(* IEC 61131-3 sources: plc-st-coding-agent/progress/evidence/f14_v14_remaining_20261113/jobs/custom_minimax-m27 (part 6) *)

(* ---- public-medium-06.raw_candidate_02.st ---- *)
FUNCTION_BLOCK FB_SlabThicknessMonitor
(*
 * ENGINEERING_CONTRACT
 * =============================================================================
 * Output/State          | Activation          | Retention            | Reset/Deactivation            | Units
 * ----------------------+---------------------+----------------------+-------------------------------+-----------------
 * THICKNESS_ALARM       | Rising edge valid   | Min 500ms hold;      | Signal invalid clears all     | BOOL
 *                       | THICKNESS_FAULT     | continues if fault   | alarm and hold state (PUB001) |
 * Alarm hold timer      | TON(IN: valid &     | TON.ET saturates at  | Signal invalid resets TON     | LTIME (≥500ms)
 *                       |   (fault OR holding))| PT=500ms            |                               |
 * Holding flag          | Fault OR holding    | Self-holds while     | Signal invalid clears         | BOOL
 *                       |                     |   fault OR timer run |                               |
 * Slab_Fault_Counter    | FALSE→TRUE valid    | Accumulates monoton  | None by task spec             | UINT
 *                       | fault transition    | (never auto-reset)   |                               |
 * Slab_Fault_History[0] | New fault entry     | Shifts [n]→[n+1]     | Power-up init to 0            | ARRAY[0..4] DINT
 *                       | writes to index 0   | (0 newest)           |                               |
 * Slab_Runtime_Accumulator| While CUTTING_RUN  | Preserved when       | None by task spec             | LTIME (accumulates)
 *                       | + valid + no fault  | conditions not met   |                               |
 * =============================================================================
 * CONTRACT_RULES [{"kind": "hold_until_reset", "output": "THICKNESS_ALARM", "set_input": "THICKNESS_FAULT", "reset_input": null}]
 *)

VAR_INPUT
    THICKNESS_FAULT        : BOOL;
    THICKNESS_SIGNAL_VALID : BOOL;
    CUTTING_RUN            : BOOL;
    FaultTimestamp         : DINT;
    CycleTime              : TIME;
END_VAR

VAR_OUTPUT
    THICKNESS_ALARM           : BOOL;
    Slab_Fault_Counter        : UINT;
    Slab_Runtime_Accumulator  : LTIME;
    Slab_Fault_History        : ARRAY[0..4] OF DINT;
END_VAR

VAR
    faultRisingEdge    : R_TRIG;
    signalValidPrev    : BOOL;
    alarmHoldTimer     : TON;
    alarmHolding       : BOOL;
    faultActive        : BOOL;
END_VAR

// ---------------------------------------------------------------------------
// Power-up initialization (first scan after instantiation)
// ---------------------------------------------------------------------------
IF NOT alarmHoldTimer.Q AND NOT faultActive AND NOT alarmHolding THEN
    Slab_Fault_Counter       := 0;
    Slab_Runtime_Accumulator := LTIME#0;
    Slab_Fault_History[0]    := 0;
    Slab_Fault_History[1]    := 0;
    Slab_Fault_History[2]    := 0;
    Slab_Fault_History[3]    := 0;
    Slab_Fault_History[4]    := 0;
END_IF;

// ---------------------------------------------------------------------------
// Detect FALSE→TRUE transition on valid fault signal
// ---------------------------------------------------------------------------
faultRisingEdge(CLK := THICKNESS_FAULT AND THICKNESS_SIGNAL_VALID);

// ---------------------------------------------------------------------------
// Handle signal-valid transitions: clear alarm/hold when signal lost (PUB001)
// ---------------------------------------------------------------------------
IF THICKNESS_SIGNAL_VALID THEN
    IF NOT signalValidPrev THEN
        // Signal just restored after being invalid
        alarmHolding  := FALSE;
        alarmHoldTimer(IN := FALSE);
        faultActive   := FALSE;
    END_IF;

    // -------------------------------------------------------------------------
    // On rising edge of valid fault: record entry and start hold
    // -------------------------------------------------------------------------
    IF faultRisingEdge.Q THEN
        // Increment counter
        Slab_Fault_Counter := Slab_Fault_Counter + UINT#1;

        // Shift history: index 3→4, 2→3, 1→2, 0→1, then write new to 0
        Slab_Fault_History[4] := Slab_Fault_History[3];
        Slab_Fault_History[3] := Slab_Fault_History[2];
        Slab_Fault_History[2] := Slab_Fault_History[1];
        Slab_Fault_History[1] := Slab_Fault_History[0];
        Slab_Fault_History[0] := FaultTimestamp;

        // Activate alarm and start 500 ms hold timer
        faultActive        := TRUE;
        alarmHolding       := TRUE;
        alarmHoldTimer(IN  := TRUE, PT := T#500ms);
    END_IF;

    // -------------------------------------------------------------------------
    // Update alarm state: hold while fault persists or timer running
    // -------------------------------------------------------------------------
    IF faultActive THEN
        // Keep timer running while fault is present
        alarmHoldTimer(IN := TRUE, PT := T#500ms);

        // Alarm stays active while fault or hold timer active
        alarmHolding := THICKNESS_FAULT OR alarmHoldTimer.Q;

        // Release hold tracking once fault clears and timer completes
        IF NOT THICKNESS_FAULT AND alarmHolding AND NOT alarmHoldTimer.Q THEN
            alarmHolding := FALSE;
        END_IF;

        // Clear fault-active flag when fault goes away (hold may continue)
        IF NOT THICKNESS_FAULT THEN
            faultActive := FALSE;
        END_IF;
    END_IF;

    // Final alarm output
    THICKNESS_ALARM := alarmHolding OR faultActive;

    // -------------------------------------------------------------------------
    // Runtime accumulation: only while cutting, signal valid, no fault
    // -------------------------------------------------------------------------
    IF CUTTING_RUN AND NOT THICKNESS_FAULT THEN
        Slab_Runtime_Accumulator := Slab_Runtime_Accumulator + TO_LTIME(CycleTime);
    END_IF;

ELSE
    // Signal invalid: clear alarm and all hold state (PUB001)
    THICKNESS_ALARM  := FALSE;
    alarmHolding     := FALSE;
    faultActive      := FALSE;
    alarmHoldTimer(IN := FALSE);
END_IF;

// ---------------------------------------------------------------------------
// Latch previous scan signal-valid state for edge detection
// ---------------------------------------------------------------------------
signalValidPrev := THICKNESS_SIGNAL_VALID;

END_FUNCTION_BLOCK

(* ---- public-medium-06.raw_candidate_03.st ---- *)
FUNCTION_BLOCK FB_SlabThicknessMonitor
(*
 * ENGINEERING_CONTRACT
 * =============================================================================
 * Output/State          | Activation          | Retention            | Reset/Deactivation            | Units
 * ----------------------+---------------------+----------------------+-------------------------------+-----------------
 * THICKNESS_ALARM       | Rising edge valid   | Min 500ms hold;      | Signal invalid clears all     | BOOL
 *                       | THICKNESS_FAULT     | continues if fault   | alarm and hold state (PUB001) |
 * Alarm hold timer      | TON(IN: valid &     | TON.ET saturates at  | Signal invalid resets TON     | LTIME (≥500ms)
 *                       |   (fault OR holding))| PT=500ms            |                               |
 * Holding flag          | Fault OR holding    | Self-holds while     | Signal invalid clears         | BOOL
 *                       |                     |   fault OR timer run |                               |
 * Slab_Fault_Counter    | FALSE→TRUE valid    | Accumulates monoton  | None by task spec             | UINT
 *                       | fault transition    | (never auto-reset)   |                               |
 * Slab_Fault_History[0] | New fault entry     | Shifts [n]→[n+1]     | Power-up init to 0            | ARRAY[0..4] DINT
 *                       | writes to index 0   | (0 newest)           |                               |
 * Slab_Runtime_Accumulator| While CUTTING_RUN  | Preserved when       | None by task spec             | LTIME (accumulates)
 *                       | + valid + no fault  | conditions not met   |                               |
 * =============================================================================
 * CONTRACT_RULES [{"kind": "hold_until_reset", "output": "THICKNESS_ALARM", "set_input": "THICKNESS_FAULT", "reset_input": null}]
 *)

VAR_INPUT
    THICKNESS_FAULT        : BOOL;
    THICKNESS_SIGNAL_VALID : BOOL;
    CUTTING_RUN            : BOOL;
    FaultTimestamp         : DINT;
    CycleTime              : TIME;
END_VAR

VAR_OUTPUT
    THICKNESS_ALARM           : BOOL;
    Slab_Fault_Counter        : UINT;
    Slab_Runtime_Accumulator  : LTIME;
    Slab_Fault_History        : ARRAY[0..4] OF DINT;
END_VAR

VAR
    faultRisingEdge    : R_TRIG;
    signalValidPrev    : BOOL;
    alarmHoldTimer     : TON;
    alarmHolding       : BOOL;
    faultActive        : BOOL;
END_VAR

// ---------------------------------------------------------------------------
// Power-up initialization (first scan after instantiation)
// ---------------------------------------------------------------------------
IF NOT alarmHoldTimer.Q AND NOT faultActive AND NOT alarmHolding THEN
    Slab_Fault_Counter       := 0;
    Slab_Runtime_Accumulator := LTIME#0ms;
    Slab_Fault_History[0]    := 0;
    Slab_Fault_History[1]    := 0;
    Slab_Fault_History[2]    := 0;
    Slab_Fault_History[3]    := 0;
    Slab_Fault_History[4]    := 0;
END_IF;

// ---------------------------------------------------------------------------
// Detect FALSE→TRUE transition on valid fault signal
// ---------------------------------------------------------------------------
faultRisingEdge(CLK := THICKNESS_FAULT AND THICKNESS_SIGNAL_VALID);

// ---------------------------------------------------------------------------
// Handle signal-valid transitions: clear alarm/hold when signal lost (PUB001)
// ---------------------------------------------------------------------------
IF THICKNESS_SIGNAL_VALID THEN
    IF NOT signalValidPrev THEN
        // Signal just restored after being invalid
        alarmHolding  := FALSE;
        alarmHoldTimer(IN := FALSE);
        faultActive   := FALSE;
    END_IF;

    // -------------------------------------------------------------------------
    // On rising edge of valid fault: record entry and start hold
    // -------------------------------------------------------------------------
    IF faultRisingEdge.Q THEN
        // Increment counter
        Slab_Fault_Counter := Slab_Fault_Counter + UINT#1;

        // Shift history: index 3→4, 2→3, 1→2, 0→1, then write new to 0
        Slab_Fault_History[4] := Slab_Fault_History[3];
        Slab_Fault_History[3] := Slab_Fault_History[2];
        Slab_Fault_History[2] := Slab_Fault_History[1];
        Slab_Fault_History[1] := Slab_Fault_History[0];
        Slab_Fault_History[0] := FaultTimestamp;

        // Activate alarm and start 500 ms hold timer
        faultActive        := TRUE;
        alarmHolding       := TRUE;
        alarmHoldTimer(IN  := TRUE, PT := T#500ms);
    END_IF;

    // -------------------------------------------------------------------------
    // Update alarm state: hold while fault persists or timer running
    // -------------------------------------------------------------------------
    IF faultActive THEN
        // Keep timer running while fault is present
        alarmHoldTimer(IN := TRUE, PT := T#500ms);

        // Alarm stays active while fault or hold timer active
        alarmHolding := THICKNESS_FAULT OR alarmHoldTimer.Q;

        // Release hold tracking once fault clears and timer completes
        IF NOT THICKNESS_FAULT AND alarmHolding AND NOT alarmHoldTimer.Q THEN
            alarmHolding := FALSE;
        END_IF;

        // Clear fault-active flag when fault goes away (hold may continue)
        IF NOT THICKNESS_FAULT THEN
            faultActive := FALSE;
        END_IF;
    END_IF;

    // Final alarm output
    THICKNESS_ALARM := alarmHolding OR faultActive;

    // -------------------------------------------------------------------------
    // Runtime accumulation: only while cutting, signal valid, no fault
    // -------------------------------------------------------------------------
    IF CUTTING_RUN AND NOT THICKNESS_FAULT THEN
        Slab_Runtime_Accumulator := Slab_Runtime_Accumulator + TO_LTIME(CycleTime);
    END_IF;

ELSE
    // Signal invalid: clear alarm and all hold state (PUB001)
    THICKNESS_ALARM  := FALSE;
    alarmHolding     := FALSE;
    faultActive      := FALSE;
    alarmHoldTimer(IN := FALSE);
END_IF;

// ---------------------------------------------------------------------------
// Latch previous scan signal-valid state for edge detection
// ---------------------------------------------------------------------------
signalValidPrev := THICKNESS_SIGNAL_VALID;

END_FUNCTION_BLOCK

(* ---- public-medium-07.candidate_01.st ---- *)
FUNCTION_BLOCK HVAC_MultiMode_Control
VAR_INPUT
    OCCUPANCY_DETECTED   : BOOL;
    ENERGY_SAVING_MODE   : BOOL;
    HVAC_MODE_SELECTOR   : INT;
END_VAR
VAR_OUTPUT
    SUPPLY_FAN_RUN       : BOOL := FALSE;
    TEMP_SETPOINT_ADJUST : INT  := 0;
END_VAR
VAR
    fan_delay_timer  : TON;
    tmp_fan_run      : BOOL := FALSE;
    tmp_adjust       : INT;
END_VAR

(* CONTRACT_RULES [] *)

(*
ENGINEERING_CONTRACT:
SUPPLY_FAN_RUN:
  - Activation: After 30s continuous occupancy without Night mode (PUB003)
  - Retention: Hold TRUE while conditions remain; reset immediately on occupancy loss or Night mode (PUB003)
  - Explicit Reset: Stop+reset when OCCUPANCY_DETECTED=FALSE OR HVAC_MODE_SELECTOR=3 (PUB003)
  - Same-scan priority: Timer starts fresh on first occupancy detection in Auto/Comfort/Economy mode
  - Boundary: TON.Q true when ET >= PT (30s); saturates at PT

TEMP_SETPOINT_ADJUST:
  - Auto(0): 0°C occupied; +3°C unoccupied with energy-saving, +2°C standard (PUB005)
  - Comfort(1): 0°C occupied; +1°C unoccupied (PUB006)
  - Economy(2): 0°C occupied; +4°C unoccupied (PUB007)
  - Night(3): +4°C regardless of occupancy (PUB008)
  - Energy-saving affects Auto mode only; units °C; clamped to ±4°C (PUB002)
*)

// --- Supply Fan Logic with 30s Delay ---
// Start delay only on first occupancy detection (timer TON resets when running with IN=FALSE)
fan_delay_timer(IN := OCCUPANCY_DETECTED AND (HVAC_MODE_SELECTOR <> 3),
                PT := T#30s);

tmp_fan_run := fan_delay_timer.Q;

// Stop immediately and reset timer if occupancy lost or Night mode selected
IF NOT OCCUPANCY_DETECTED OR (HVAC_MODE_SELECTOR = 3) THEN
    tmp_fan_run := FALSE;
    fan_delay_timer(IN := FALSE);
END_IF;

SUPPLY_FAN_RUN := tmp_fan_run;

// --- Temperature Setpoint Adjustment ---
CASE HVAC_MODE_SELECTOR OF
    0:  // Auto mode
        IF OCCUPANCY_DETECTED THEN
            tmp_adjust := 0;
        ELSE
            IF ENERGY_SAVING_MODE THEN
                tmp_adjust := 3;  // +3°C energy saving
            ELSE
                tmp_adjust := 2;  // +2°C standard
            END_IF;
        END_IF;

    1:  // Comfort mode
        IF OCCUPANCY_DETECTED THEN
            tmp_adjust := 0;
        ELSE
            tmp_adjust := 1;
        END_IF;

    2:  // Economy mode
        IF OCCUPANCY_DETECTED THEN
            tmp_adjust := 0;
        ELSE
            tmp_adjust := 4;
        END_IF;

    3:  // Night mode
        tmp_adjust := 4;

    ELSE
        tmp_adjust := 0;
END_CASE;

// Clamp to ±4°C per PUB002
IF tmp_adjust > 4 THEN
    tmp_adjust := 4;
ELSIF tmp_adjust < -4 THEN
    tmp_adjust := -4;
END_IF;

TEMP_SETPOINT_ADJUST := tmp_adjust;

END_FUNCTION_BLOCK

(* ---- public-medium-07.raw_candidate_01.st ---- *)
FUNCTION_BLOCK HVAC_MultiMode_Control
VAR_INPUT
    OCCUPANCY_DETECTED   : BOOL;
    ENERGY_SAVING_MODE   : BOOL;
    HVAC_MODE_SELECTOR   : INT;
END_VAR
VAR_OUTPUT
    SUPPLY_FAN_RUN       : BOOL := FALSE;
    TEMP_SETPOINT_ADJUST : INT  := 0;
END_VAR
VAR
    fan_delay_timer  : TON;
    tmp_fan_run      : BOOL := FALSE;
    tmp_adjust       : INT;
END_VAR

(* CONTRACT_RULES [] *)

(*
ENGINEERING_CONTRACT:
SUPPLY_FAN_RUN:
  - Activation: After 30s continuous occupancy without Night mode (PUB003)
  - Retention: Hold TRUE while conditions remain; reset immediately on occupancy loss or Night mode (PUB003)
  - Explicit Reset: Stop+reset when OCCUPANCY_DETECTED=FALSE OR HVAC_MODE_SELECTOR=3 (PUB003)
  - Same-scan priority: Timer starts fresh on first occupancy detection in Auto/Comfort/Economy mode
  - Boundary: TON.Q true when ET >= PT (30s); saturates at PT

TEMP_SETPOINT_ADJUST:
  - Auto(0): 0°C occupied; +3°C unoccupied with energy-saving, +2°C standard (PUB005)
  - Comfort(1): 0°C occupied; +1°C unoccupied (PUB006)
  - Economy(2): 0°C occupied; +4°C unoccupied (PUB007)
  - Night(3): +4°C regardless of occupancy (PUB008)
  - Energy-saving affects Auto mode only; units °C; clamped to ±4°C (PUB002)
*)

// --- Supply Fan Logic with 30s Delay ---
// Start delay only on first occupancy detection (timer TON resets when running with IN=FALSE)
fan_delay_timer(IN := OCCUPANCY_DETECTED AND (HVAC_MODE_SELECTOR <> 3),
                PT := T#30s);

tmp_fan_run := fan_delay_timer.Q;

// Stop immediately and reset timer if occupancy lost or Night mode selected
IF NOT OCCUPANCY_DETECTED OR (HVAC_MODE_SELECTOR = 3) THEN
    tmp_fan_run := FALSE;
    fan_delay_timer(IN := FALSE);
END_IF;

SUPPLY_FAN_RUN := tmp_fan_run;

// --- Temperature Setpoint Adjustment ---
CASE HVAC_MODE_SELECTOR OF
    0:  // Auto mode
        IF OCCUPANCY_DETECTED THEN
            tmp_adjust := 0;
        ELSE
            IF ENERGY_SAVING_MODE THEN
                tmp_adjust := 3;  // +3°C energy saving
            ELSE
                tmp_adjust := 2;  // +2°C standard
            END_IF;
        END_IF;

    1:  // Comfort mode
        IF OCCUPANCY_DETECTED THEN
            tmp_adjust := 0;
        ELSE
            tmp_adjust := 1;
        END_IF;

    2:  // Economy mode
        IF OCCUPANCY_DETECTED THEN
            tmp_adjust := 0;
        ELSE
            tmp_adjust := 4;
        END_IF;

    3:  // Night mode
        tmp_adjust := 4;

    ELSE
        tmp_adjust := 0;
END_CASE;

// Clamp to ±4°C per PUB002
IF tmp_adjust > 4 THEN
    tmp_adjust := 4;
ELSIF tmp_adjust < -4 THEN
    tmp_adjust := -4;
END_IF;

TEMP_SETPOINT_ADJUST := tmp_adjust;

END_FUNCTION_BLOCK

(* ---- public-medium-08.candidate_01.st ---- *)
FUNCTION_BLOCK FB_IPv4Parse
VAR_INPUT
    ipText : STRING(254);
END_VAR
VAR_OUTPUT
    ipValue : UDINT;
END_VAR
VAR
    tmp_dot1 : INT;
    tmp_dot2 : INT;
    tmp_dot3 : INT;
    tmp_seg1 : STRING(4);
    tmp_seg2 : STRING(4);
    tmp_seg3 : STRING(4);
    tmp_seg4 : STRING(4);
    tmp_val1 : UDINT;
    tmp_val2 : UDINT;
    tmp_val3 : UDINT;
    tmp_val4 : UDINT;
    tmp_valid : BOOL;
    tmp_i : INT;
    tmp_ch : BYTE;
END_VAR
(* ENGINEERING_CONTRACT
 * Parse dotted-decimal IPv4 string to 32-bit network-order UDINT.
 * Input:  ipText (STRING(254)) - dotted-decimal address
 * Output: ipValue (UDINT) - 32-bit value, network byte order; 0 if invalid
 *
 * PUB001: Parse ipText for exactly 4 decimal-digit segments separated by 3 periods
 * PUB002: Each segment value must be 0-255 inclusive
 * PUB003: Network byte order: seg1=MSB<<24, seg2<<16, seg3<<8, seg4=LSB
 * PUB004: Invalid input (wrong count, nondigit, OOR, empty segment) → ipValue=0
 *         Note: Valid address 0.0.0.0 also produces 0 per spec.
 *
 * Contract behavior: Pure combinational, no latches, no state retention.
 * Output ipValue is defined every scan from current ipText.
 *)

ipValue := 0;
tmp_valid := TRUE;

tmp_dot1 := FIND(ipText, '.');
IF tmp_dot1 < 2 OR tmp_dot1 >= LEN(ipText) THEN
    tmp_valid := FALSE;
END_IF;

IF tmp_valid THEN
    tmp_dot2 := FIND(MID(ipText, LEN(ipText) - tmp_dot1, tmp_dot1 + 1), '.');
    IF tmp_dot2 < 2 OR tmp_dot2 >= (LEN(ipText) - tmp_dot1) THEN
        tmp_valid := FALSE;
    END_IF;
END_IF;

IF tmp_valid THEN
    tmp_dot3 := FIND(MID(ipText, LEN(ipText) - (tmp_dot1 + tmp_dot2), tmp_dot1 + tmp_dot2 + 1), '.');
    IF tmp_dot3 < 2 THEN
        tmp_valid := FALSE;
    END_IF;
END_IF;

IF tmp_valid THEN
    tmp_seg1 := LEFT(ipText, tmp_dot1 - 1);
    tmp_seg2 := MID(ipText, tmp_dot2 - 1, tmp_dot1 + 1);
    tmp_seg3 := MID(ipText, tmp_dot3 - 1, tmp_dot1 + tmp_dot2 + 1);
    tmp_seg4 := MID(ipText, LEN(ipText) - (tmp_dot1 + tmp_dot2 + tmp_dot3), tmp_dot1 + tmp_dot2 + tmp_dot3 + 1);

    // Validate segment 1
    IF LEN(tmp_seg1) < 1 OR LEN(tmp_seg1) > 3 THEN
        tmp_valid := FALSE;
    ELSE
        tmp_val1 := 0;
        FOR tmp_i := 1 TO LEN(tmp_seg1) DO
            tmp_ch := MID(tmp_seg1, 1, tmp_i);
            IF tmp_ch < 48 OR tmp_ch > 57 THEN
                tmp_valid := FALSE;
                EXIT;
            END_IF;
            tmp_val1 := tmp_val1 * 10 + TO_UDINT(tmp_ch - 48);
        END_FOR;
        IF tmp_val1 > 255 THEN
            tmp_valid := FALSE;
        END_IF;
    END_IF;

    // Validate segment 2
    IF tmp_valid AND (LEN(tmp_seg2) < 1 OR LEN(tmp_seg2) > 3) THEN
        tmp_valid := FALSE;
    END_IF;

    IF tmp_valid THEN
        tmp_val2 := 0;
        FOR tmp_i := 1 TO LEN(tmp_seg2) DO
            tmp_ch := MID(tmp_seg2, 1, tmp_i);
            IF tmp_ch < 48 OR tmp_ch > 57 THEN
                tmp_valid := FALSE;
                EXIT;
            END_IF;
            tmp_val2 := tmp_val2 * 10 + TO_UDINT(tmp_ch - 48);
        END_FOR;
        IF tmp_val2 > 255 THEN
            tmp_valid := FALSE;
        END_IF;
    END_IF;

    // Validate segment 3
    IF tmp_valid AND (LEN(tmp_seg3) < 1 OR LEN(tmp_seg3) > 3) THEN
        tmp_valid := FALSE;
    END_IF;

    IF tmp_valid THEN
        tmp_val3 := 0;
        FOR tmp_i := 1 TO LEN(tmp_seg3) DO
            tmp_ch := MID(tmp_seg3, 1, tmp_i);
            IF tmp_ch < 48 OR tmp_ch > 57 THEN
                tmp_valid := FALSE;
                EXIT;
            END_IF;
            tmp_val3 := tmp_val3 * 10 + TO_UDINT(tmp_ch - 48);
        END_FOR;
        IF tmp_val3 > 255 THEN
            tmp_valid := FALSE;
        END_IF;
    END_IF;

    // Validate segment 4
    IF tmp_valid AND (LEN(tmp_seg4) < 1 OR LEN(tmp_seg4) > 3) THEN
        tmp_valid := FALSE;
    END_IF;

    IF tmp_valid THEN
        tmp_val4 := 0;
        FOR tmp_i := 1 TO LEN(tmp_seg4) DO
            tmp_ch := MID(tmp_seg4, 1, tmp_i);
            IF tmp_ch < 48 OR tmp_ch > 57 THEN
                tmp_valid := FALSE;
                EXIT;
            END_IF;
            tmp_val4 := tmp_val4 * 10 + TO_UDINT(tmp_ch - 48);
        END_FOR;
        IF tmp_val4 > 255 THEN
            tmp_valid := FALSE;
        END_IF;
    END_IF;
END_IF;

IF tmp_valid THEN
    ipValue := SHL(tmp_val1, 24) OR SHL(tmp_val2, 16) OR SHL(tmp_val3, 8) OR tmp_val4;
END_IF;

END_FUNCTION_BLOCK
(* CONTRACT_RULES [] *)

(* ---- public-medium-08.candidate_03.st ---- *)
FUNCTION_BLOCK FB_IPv4Parse
VAR_INPUT
    ipText : STRING(254);
END_VAR
VAR_OUTPUT
    ipValue : UDINT;
END_VAR
VAR
    tmp_dot1 : INT;
    tmp_dot2 : INT;
    tmp_dot3 : INT;
    tmp_seg1 : STRING(4);
    tmp_seg2 : STRING(4);
    tmp_seg3 : STRING(4);
    tmp_seg4 : STRING(4);
    tmp_val1 : UDINT;
    tmp_val2 : UDINT;
    tmp_val3 : UDINT;
    tmp_val4 : UDINT;
    tmp_valid : BOOL;
    tmp_i : INT;
    tmp_ch : BYTE;
END_VAR
(* ENGINEERING_CONTRACT
 * Parse dotted-decimal IPv4 string to 32-bit network-order UDINT.
 * Input:  ipText (STRING(254)) - dotted-decimal address
 * Output: ipValue (UDINT) - 32-bit value, network byte order; 0 if invalid
 *
 * PUB001: Parse ipText for exactly 4 decimal-digit segments separated by 3 periods
 * PUB002: Each segment value must be 0-255 inclusive
 * PUB003: Network byte order: seg1=MSB<<24, seg2<<16, seg3<<8, seg4=LSB
 * PUB004: Invalid input (wrong count, nondigit, OOR, empty segment) → ipValue=0
 *         Note: Valid address 0.0.0.0 also produces 0 per spec.
 *
 * Contract behavior: Pure combinational, no latches, no state retention.
 * Output ipValue is defined every scan from current ipText.
 *)

ipValue := 0;
tmp_valid := TRUE;

tmp_dot1 := FIND(ipText, '.');
IF tmp_dot1 < 2 OR tmp_dot1 >= LEN(ipText) THEN
    tmp_valid := FALSE;
END_IF;

IF tmp_valid THEN
    tmp_dot2 := FIND(MID(ipText, LEN(ipText) - tmp_dot1, tmp_dot1 + 1), '.');
    IF tmp_dot2 < 2 OR tmp_dot2 >= (LEN(ipText) - tmp_dot1) THEN
        tmp_valid := FALSE;
    END_IF;
END_IF;

IF tmp_valid THEN
    tmp_dot3 := FIND(MID(ipText, LEN(ipText) - (tmp_dot1 + tmp_dot2), tmp_dot1 + tmp_dot2 + 1), '.');
    IF tmp_dot3 < 2 THEN
        tmp_valid := FALSE;
    END_IF;
END_IF;

IF tmp_valid THEN
    tmp_seg1 := LEFT(ipText, tmp_dot1 - 1);
    tmp_seg2 := MID(ipText, tmp_dot2 - 1, tmp_dot1 + 1);
    tmp_seg3 := MID(ipText, tmp_dot3 - 1, tmp_dot1 + tmp_dot2 + 1);
    tmp_seg4 := MID(ipText, LEN(ipText) - (tmp_dot1 + tmp_dot2 + tmp_dot3), tmp_dot1 + tmp_dot2 + tmp_dot3 + 1);

    // Validate segment 1
    IF LEN(tmp_seg1) < 1 OR LEN(tmp_seg1) > 3 THEN
        tmp_valid := FALSE;
    ELSE
        tmp_val1 := 0;
        FOR tmp_i := 1 TO LEN(tmp_seg1) DO
            tmp_ch := ipText[tmp_i];
            IF tmp_ch < 48 OR tmp_ch > 57 THEN
                tmp_valid := FALSE;
                EXIT;
            END_IF;
            tmp_val1 := tmp_val1 * 10 + TO_UDINT(tmp_ch - 48);
        END_FOR;
        IF tmp_val1 > 255 THEN
            tmp_valid := FALSE;
        END_IF;
    END_IF;

    // Validate segment 2
    IF tmp_valid AND (LEN(tmp_seg2) < 1 OR LEN(tmp_seg2) > 3) THEN
        tmp_valid := FALSE;
    END_IF;

    IF tmp_valid THEN
        tmp_val2 := 0;
        FOR tmp_i := 1 TO LEN(tmp_seg2) DO
            tmp_ch := ipText[tmp_dot1 + tmp_dot2 + tmp_i];
            IF tmp_ch < 48 OR tmp_ch > 57 THEN
                tmp_valid := FALSE;
                EXIT;
            END_IF;
            tmp_val2 := tmp_val2 * 10 + TO_UDINT(tmp_ch - 48);
        END_FOR;
        IF tmp_val2 > 255 THEN
            tmp_valid := FALSE;
        END_IF;
    END_IF;

    // Validate segment 3
    IF tmp_valid AND (LEN(tmp_seg3) < 1 OR LEN(tmp_seg3) > 3) THEN
        tmp_valid := FALSE;
    END_IF;

    IF tmp_valid THEN
        tmp_val3 := 0;
        FOR tmp_i := 1 TO LEN(tmp_seg3) DO
            tmp_ch := ipText[tmp_dot1 + tmp_dot2 + tmp_dot3 + tmp_i];
            IF tmp_ch < 48 OR tmp_ch > 57 THEN
                tmp_valid := FALSE;
                EXIT;
            END_IF;
            tmp_val3 := tmp_val3 * 10 + TO_UDINT(tmp_ch - 48);
        END_FOR;
        IF tmp_val3 > 255 THEN
            tmp_valid := FALSE;
        END_IF;
    END_IF;

    // Validate segment 4
    IF tmp_valid AND (LEN(tmp_seg4) < 1 OR LEN(tmp_seg4) > 3) THEN
        tmp_valid := FALSE;
    END_IF;

    IF tmp_valid THEN
        tmp_val4 := 0;
        FOR tmp_i := 1 TO LEN(tmp_seg4) DO
            tmp_ch := ipText[tmp_dot1 + tmp_dot2 + tmp_dot3 + tmp_i];
            IF tmp_ch < 48 OR tmp_ch > 57 THEN
                tmp_valid := FALSE;
                EXIT;
            END_IF;
            tmp_val4 := tmp_val4 * 10 + TO_UDINT(tmp_ch - 48);
        END_FOR;
        IF tmp_val4 > 255 THEN
            tmp_valid := FALSE;
        END_IF;
    END_IF;
END_IF;

IF tmp_valid THEN
    ipValue := SHL(tmp_val1, 24) OR SHL(tmp_val2, 16) OR SHL(tmp_val3, 8) OR tmp_val4;
END_IF;

END_FUNCTION_BLOCK
(* CONTRACT_RULES [] *)

(* ---- public-medium-08.patch_base_02.st ---- *)
FUNCTION_BLOCK FB_IPv4Parse
VAR_INPUT
    ipText : STRING(254);
END_VAR
VAR_OUTPUT
    ipValue : UDINT;
END_VAR
VAR
    tmp_dot1 : INT;
    tmp_dot2 : INT;
    tmp_dot3 : INT;
    tmp_seg1 : STRING(4);
    tmp_seg2 : STRING(4);
    tmp_seg3 : STRING(4);
    tmp_seg4 : STRING(4);
    tmp_val1 : UDINT;
    tmp_val2 : UDINT;
    tmp_val3 : UDINT;
    tmp_val4 : UDINT;
    tmp_valid : BOOL;
    tmp_i : INT;
    tmp_ch : BYTE;
END_VAR
(* ENGINEERING_CONTRACT
 * Parse dotted-decimal IPv4 string to 32-bit network-order UDINT.
 * Input:  ipText (STRING(254)) - dotted-decimal address
 * Output: ipValue (UDINT) - 32-bit value, network byte order; 0 if invalid
 *
 * PUB001: Parse ipText for exactly 4 decimal-digit segments separated by 3 periods
 * PUB002: Each segment value must be 0-255 inclusive
 * PUB003: Network byte order: seg1=MSB<<24, seg2<<16, seg3<<8, seg4=LSB
 * PUB004: Invalid input (wrong count, nondigit, OOR, empty segment) → ipValue=0
 *         Note: Valid address 0.0.0.0 also produces 0 per spec.
 *
 * Contract behavior: Pure combinational, no latches, no state retention.
 * Output ipValue is defined every scan from current ipText.
 *)

ipValue := 0;
tmp_valid := TRUE;

tmp_dot1 := FIND(ipText, '.');
IF tmp_dot1 < 2 OR tmp_dot1 >= LEN(ipText) THEN
    tmp_valid := FALSE;
END_IF;

IF tmp_valid THEN
    tmp_dot2 := FIND(MID(ipText, LEN(ipText) - tmp_dot1, tmp_dot1 + 1), '.');
    IF tmp_dot2 < 2 OR tmp_dot2 >= (LEN(ipText) - tmp_dot1) THEN
        tmp_valid := FALSE;
    END_IF;
END_IF;

IF tmp_valid THEN
    tmp_dot3 := FIND(MID(ipText, LEN(ipText) - (tmp_dot1 + tmp_dot2), tmp_dot1 + tmp_dot2 + 1), '.');
    IF tmp_dot3 < 2 THEN
        tmp_valid := FALSE;
    END_IF;
END_IF;

IF tmp_valid THEN
    tmp_seg1 := LEFT(ipText, tmp_dot1 - 1);
    tmp_seg2 := MID(ipText, tmp_dot2 - 1, tmp_dot1 + 1);
    tmp_seg3 := MID(ipText, tmp_dot3 - 1, tmp_dot1 + tmp_dot2 + 1);
    tmp_seg4 := MID(ipText, LEN(ipText) - (tmp_dot1 + tmp_dot2 + tmp_dot3), tmp_dot1 + tmp_dot2 + tmp_dot3 + 1);

    // Validate segment 1
    IF LEN(tmp_seg1) < 1 OR LEN(tmp_seg1) > 3 THEN
        tmp_valid := FALSE;
    ELSE
        tmp_val1 := 0;
        FOR tmp_i := 1 TO LEN(tmp_seg1) DO
            tmp_ch := MID(tmp_seg1, 1, tmp_i);
            IF tmp_ch < 48 OR tmp_ch > 57 THEN
                tmp_valid := FALSE;
                EXIT;
            END_IF;
            tmp_val1 := tmp_val1 * 10 + TO_UDINT(tmp_ch - 48);
        END_FOR;
        IF tmp_val1 > 255 THEN
            tmp_valid := FALSE;
        END_IF;
    END_IF;

    // Validate segment 2
    IF tmp_valid AND (LEN(tmp_seg2) < 1 OR LEN(tmp_seg2) > 3) THEN
        tmp_valid := FALSE;
    END_IF;

    IF tmp_valid THEN
        tmp_val2 := 0;
        FOR tmp_i := 1 TO LEN(tmp_seg2) DO
            tmp_ch := MID(tmp_seg2, 1, tmp_i);
            IF tmp_ch < 48 OR tmp_ch > 57 THEN
                tmp_valid := FALSE;
                EXIT;
            END_IF;
            tmp_val2 := tmp_val2 * 10 + TO_UDINT(tmp_ch - 48);
        END_FOR;
        IF tmp_val2 > 255 THEN
            tmp_valid := FALSE;
        END_IF;
    END_IF;

    // Validate segment 3
    IF tmp_valid AND (LEN(tmp_seg3) < 1 OR LEN(tmp_seg3) > 3) THEN
        tmp_valid := FALSE;
    END_IF;

    IF tmp_valid THEN
        tmp_val3 := 0;
        FOR tmp_i := 1 TO LEN(tmp_seg3) DO
            tmp_ch := MID(tmp_seg3, 1, tmp_i);
            IF tmp_ch < 48 OR tmp_ch > 57 THEN
                tmp_valid := FALSE;
                EXIT;
            END_IF;
            tmp_val3 := tmp_val3 * 10 + TO_UDINT(tmp_ch - 48);
        END_FOR;
        IF tmp_val3 > 255 THEN
            tmp_valid := FALSE;
        END_IF;
    END_IF;

    // Validate segment 4
    IF tmp_valid AND (LEN(tmp_seg4) < 1 OR LEN(tmp_seg4) > 3) THEN
        tmp_valid := FALSE;
    END_IF;

    IF tmp_valid THEN
        tmp_val4 := 0;
        FOR tmp_i := 1 TO LEN(tmp_seg4) DO
            tmp_ch := MID(tmp_seg4, 1, tmp_i);
            IF tmp_ch < 48 OR tmp_ch > 57 THEN
                tmp_valid := FALSE;
                EXIT;
            END_IF;
            tmp_val4 := tmp_val4 * 10 + TO_UDINT(tmp_ch - 48);
        END_FOR;
        IF tmp_val4 > 255 THEN
            tmp_valid := FALSE;
        END_IF;
    END_IF;
END_IF;

IF tmp_valid THEN
    ipValue := SHL(tmp_val1, 24) OR SHL(tmp_val2, 16) OR SHL(tmp_val3, 8) OR tmp_val4;
END_IF;

END_FUNCTION_BLOCK
(* CONTRACT_RULES [] *)

(* ---- public-medium-08.patch_base_03.st ---- *)
FUNCTION_BLOCK FB_IPv4Parse
VAR_INPUT
    ipText : STRING(254);
END_VAR
VAR_OUTPUT
    ipValue : UDINT;
END_VAR
VAR
    tmp_dot1 : INT;
    tmp_dot2 : INT;
    tmp_dot3 : INT;
    tmp_seg1 : STRING(4);
    tmp_seg2 : STRING(4);
    tmp_seg3 : STRING(4);
    tmp_seg4 : STRING(4);
    tmp_val1 : UDINT;
    tmp_val2 : UDINT;
    tmp_val3 : UDINT;
    tmp_val4 : UDINT;
    tmp_valid : BOOL;
    tmp_i : INT;
    tmp_ch : BYTE;
END_VAR
(* ENGINEERING_CONTRACT
 * Parse dotted-decimal IPv4 string to 32-bit network-order UDINT.
 * Input:  ipText (STRING(254)) - dotted-decimal address
 * Output: ipValue (UDINT) - 32-bit value, network byte order; 0 if invalid
 *
 * PUB001: Parse ipText for exactly 4 decimal-digit segments separated by 3 periods
 * PUB002: Each segment value must be 0-255 inclusive
 * PUB003: Network byte order: seg1=MSB<<24, seg2<<16, seg3<<8, seg4=LSB
 * PUB004: Invalid input (wrong count, nondigit, OOR, empty segment) → ipValue=0
 *         Note: Valid address 0.0.0.0 also produces 0 per spec.
 *
 * Contract behavior: Pure combinational, no latches, no state retention.
 * Output ipValue is defined every scan from current ipText.
 *)

ipValue := 0;
tmp_valid := TRUE;

tmp_dot1 := FIND(ipText, '.');
IF tmp_dot1 < 2 OR tmp_dot1 >= LEN(ipText) THEN
    tmp_valid := FALSE;
END_IF;

IF tmp_valid THEN
    tmp_dot2 := FIND(MID(ipText, LEN(ipText) - tmp_dot1, tmp_dot1 + 1), '.');
    IF tmp_dot2 < 2 OR tmp_dot2 >= (LEN(ipText) - tmp_dot1) THEN
        tmp_valid := FALSE;
    END_IF;
END_IF;

IF tmp_valid THEN
    tmp_dot3 := FIND(MID(ipText, LEN(ipText) - (tmp_dot1 + tmp_dot2), tmp_dot1 + tmp_dot2 + 1), '.');
    IF tmp_dot3 < 2 THEN
        tmp_valid := FALSE;
    END_IF;
END_IF;

IF tmp_valid THEN
    tmp_seg1 := LEFT(ipText, tmp_dot1 - 1);
    tmp_seg2 := MID(ipText, tmp_dot2 - 1, tmp_dot1 + 1);
    tmp_seg3 := MID(ipText, tmp_dot3 - 1, tmp_dot1 + tmp_dot2 + 1);
    tmp_seg4 := MID(ipText, LEN(ipText) - (tmp_dot1 + tmp_dot2 + tmp_dot3), tmp_dot1 + tmp_dot2 + tmp_dot3 + 1);

    // Validate segment 1
    IF LEN(tmp_seg1) < 1 OR LEN(tmp_seg1) > 3 THEN
        tmp_valid := FALSE;
    ELSE
        tmp_val1 := 0;
        FOR tmp_i := 1 TO LEN(tmp_seg1) DO
            tmp_ch := MID(tmp_seg1, 1, tmp_i);
            IF tmp_ch < 48 OR tmp_ch > 57 THEN
                tmp_valid := FALSE;
                EXIT;
            END_IF;
            tmp_val1 := tmp_val1 * 10 + TO_UDINT(tmp_ch - 48);
        END_FOR;
        IF tmp_val1 > 255 THEN
            tmp_valid := FALSE;
        END_IF;
    END_IF;

    // Validate segment 2
    IF tmp_valid AND (LEN(tmp_seg2) < 1 OR LEN(tmp_seg2) > 3) THEN
        tmp_valid := FALSE;
    END_IF;

    IF tmp_valid THEN
        tmp_val2 := 0;
        FOR tmp_i := 1 TO LEN(tmp_seg2) DO
            tmp_ch := MID(tmp_seg2, 1, tmp_i);
            IF tmp_ch < 48 OR tmp_ch > 57 THEN
                tmp_valid := FALSE;
                EXIT;
            END_IF;
            tmp_val2 := tmp_val2 * 10 + TO_UDINT(tmp_ch - 48);
        END_FOR;
        IF tmp_val2 > 255 THEN
            tmp_valid := FALSE;
        END_IF;
    END_IF;

    // Validate segment 3
    IF tmp_valid AND (LEN(tmp_seg3) < 1 OR LEN(tmp_seg3) > 3) THEN
        tmp_valid := FALSE;
    END_IF;

    IF tmp_valid THEN
        tmp_val3 := 0;
        FOR tmp_i := 1 TO LEN(tmp_seg3) DO
            tmp_ch := MID(tmp_seg3, 1, tmp_i);
            IF tmp_ch < 48 OR tmp_ch > 57 THEN
                tmp_valid := FALSE;
                EXIT;
            END_IF;
            tmp_val3 := tmp_val3 * 10 + TO_UDINT(tmp_ch - 48);
        END_FOR;
        IF tmp_val3 > 255 THEN
            tmp_valid := FALSE;
        END_IF;
    END_IF;

    // Validate segment 4
    IF tmp_valid AND (LEN(tmp_seg4) < 1 OR LEN(tmp_seg4) > 3) THEN
        tmp_valid := FALSE;
    END_IF;

    IF tmp_valid THEN
        tmp_val4 := 0;
        FOR tmp_i := 1 TO LEN(tmp_seg4) DO
            tmp_ch := MID(tmp_seg4, 1, tmp_i);
            IF tmp_ch < 48 OR tmp_ch > 57 THEN
                tmp_valid := FALSE;
                EXIT;
            END_IF;
            tmp_val4 := tmp_val4 * 10 + TO_UDINT(tmp_ch - 48);
        END_FOR;
        IF tmp_val4 > 255 THEN
            tmp_valid := FALSE;
        END_IF;
    END_IF;
END_IF;

IF tmp_valid THEN
    ipValue := SHL(tmp_val1, 24) OR SHL(tmp_val2, 16) OR SHL(tmp_val3, 8) OR tmp_val4;
END_IF;

END_FUNCTION_BLOCK
(* CONTRACT_RULES [] *)

(* ---- public-medium-08.patch_base_04.st ---- *)
FUNCTION_BLOCK FB_IPv4Parse
VAR_INPUT
    ipText : STRING(254);
END_VAR
VAR_OUTPUT
    ipValue : UDINT;
END_VAR
VAR
    tmp_dot1 : INT;
    tmp_dot2 : INT;
    tmp_dot3 : INT;
    tmp_seg1 : STRING(4);
    tmp_seg2 : STRING(4);
    tmp_seg3 : STRING(4);
    tmp_seg4 : STRING(4);
    tmp_val1 : UDINT;
    tmp_val2 : UDINT;
    tmp_val3 : UDINT;
    tmp_val4 : UDINT;
    tmp_valid : BOOL;
    tmp_i : INT;
    tmp_ch : BYTE;
END_VAR
(* ENGINEERING_CONTRACT
 * Parse dotted-decimal IPv4 string to 32-bit network-order UDINT.
 * Input:  ipText (STRING(254)) - dotted-decimal address
 * Output: ipValue (UDINT) - 32-bit value, network byte order; 0 if invalid
 *
 * PUB001: Parse ipText for exactly 4 decimal-digit segments separated by 3 periods
 * PUB002: Each segment value must be 0-255 inclusive
 * PUB003: Network byte order: seg1=MSB<<24, seg2<<16, seg3<<8, seg4=LSB
 * PUB004: Invalid input (wrong count, nondigit, OOR, empty segment) → ipValue=0
 *         Note: Valid address 0.0.0.0 also produces 0 per spec.
 *
 * Contract behavior: Pure combinational, no latches, no state retention.
 * Output ipValue is defined every scan from current ipText.
 *)

ipValue := 0;
tmp_valid := TRUE;

tmp_dot1 := FIND(ipText, '.');
IF tmp_dot1 < 2 OR tmp_dot1 >= LEN(ipText) THEN
    tmp_valid := FALSE;
END_IF;

IF tmp_valid THEN
    tmp_dot2 := FIND(MID(ipText, LEN(ipText) - tmp_dot1, tmp_dot1 + 1), '.');
    IF tmp_dot2 < 2 OR tmp_dot2 >= (LEN(ipText) - tmp_dot1) THEN
        tmp_valid := FALSE;
    END_IF;
END_IF;

IF tmp_valid THEN
    tmp_dot3 := FIND(MID(ipText, LEN(ipText) - (tmp_dot1 + tmp_dot2), tmp_dot1 + tmp_dot2 + 1), '.');
    IF tmp_dot3 < 2 THEN
        tmp_valid := FALSE;
    END_IF;
END_IF;

IF tmp_valid THEN
    tmp_seg1 := LEFT(ipText, tmp_dot1 - 1);
    tmp_seg2 := MID(ipText, tmp_dot2 - 1, tmp_dot1 + 1);
    tmp_seg3 := MID(ipText, tmp_dot3 - 1, tmp_dot1 + tmp_dot2 + 1);
    tmp_seg4 := MID(ipText, LEN(ipText) - (tmp_dot1 + tmp_dot2 + tmp_dot3), tmp_dot1 + tmp_dot2 + tmp_dot3 + 1);

    // Validate segment 1
    IF LEN(tmp_seg1) < 1 OR LEN(tmp_seg1) > 3 THEN
        tmp_valid := FALSE;
    ELSE
        tmp_val1 := 0;
        FOR tmp_i := 1 TO LEN(tmp_seg1) DO
            tmp_ch := ipText[tmp_i];
            IF tmp_ch < 48 OR tmp_ch > 57 THEN
                tmp_valid := FALSE;
                EXIT;
            END_IF;
            tmp_val1 := tmp_val1 * 10 + TO_UDINT(tmp_ch - 48);
        END_FOR;
        IF tmp_val1 > 255 THEN
            tmp_valid := FALSE;
        END_IF;
    END_IF;

    // Validate segment 2
    IF tmp_valid AND (LEN(tmp_seg2) < 1 OR LEN(tmp_seg2) > 3) THEN
        tmp_valid := FALSE;
    END_IF;

    IF tmp_valid THEN
        tmp_val2 := 0;
        FOR tmp_i := 1 TO LEN(tmp_seg2) DO
            tmp_ch := ipText[tmp_dot1 + tmp_dot2 + tmp_i];
            IF tmp_ch < 48 OR tmp_ch > 57 THEN
                tmp_valid := FALSE;
                EXIT;
            END_IF;
            tmp_val2 := tmp_val2 * 10 + TO_UDINT(tmp_ch - 48);
        END_FOR;
        IF tmp_val2 > 255 THEN
            tmp_valid := FALSE;
        END_IF;
    END_IF;

    // Validate segment 3
    IF tmp_valid AND (LEN(tmp_seg3) < 1 OR LEN(tmp_seg3) > 3) THEN
        tmp_valid := FALSE;
    END_IF;

    IF tmp_valid THEN
        tmp_val3 := 0;
        FOR tmp_i := 1 TO LEN(tmp_seg3) DO
            tmp_ch := ipText[tmp_dot1 + tmp_dot2 + tmp_dot3 + tmp_i];
            IF tmp_ch < 48 OR tmp_ch > 57 THEN
                tmp_valid := FALSE;
                EXIT;
            END_IF;
            tmp_val3 := tmp_val3 * 10 + TO_UDINT(tmp_ch - 48);
        END_FOR;
        IF tmp_val3 > 255 THEN
            tmp_valid := FALSE;
        END_IF;
    END_IF;

    // Validate segment 4
    IF tmp_valid AND (LEN(tmp_seg4) < 1 OR LEN(tmp_seg4) > 3) THEN
        tmp_valid := FALSE;
    END_IF;

    IF tmp_valid THEN
        tmp_val4 := 0;
        FOR tmp_i := 1 TO LEN(tmp_seg4) DO
            tmp_ch := ipText[tmp_dot1 + tmp_dot2 + tmp_dot3 + tmp_i];
            IF tmp_ch < 48 OR tmp_ch > 57 THEN
                tmp_valid := FALSE;
                EXIT;
            END_IF;
            tmp_val4 := tmp_val4 * 10 + TO_UDINT(tmp_ch - 48);
        END_FOR;
        IF tmp_val4 > 255 THEN
            tmp_valid := FALSE;
        END_IF;
    END_IF;
END_IF;

IF tmp_valid THEN
    ipValue := SHL(tmp_val1, 24) OR SHL(tmp_val2, 16) OR SHL(tmp_val3, 8) OR tmp_val4;
END_IF;

END_FUNCTION_BLOCK
(* CONTRACT_RULES [] *)

(* ---- public-medium-08.raw_candidate_01.st ---- *)
FUNCTION_BLOCK FB_IPv4Parse
VAR_INPUT
    ipText : STRING(254);
END_VAR
VAR_OUTPUT
    ipValue : UDINT;
END_VAR
VAR
    tmp_dot1 : INT;
    tmp_dot2 : INT;
    tmp_dot3 : INT;
    tmp_seg1 : STRING(4);
    tmp_seg2 : STRING(4);
    tmp_seg3 : STRING(4);
    tmp_seg4 : STRING(4);
    tmp_val1 : UDINT;
    tmp_val2 : UDINT;
    tmp_val3 : UDINT;
    tmp_val4 : UDINT;
    tmp_valid : BOOL;
    tmp_i : INT;
    tmp_ch : BYTE;
END_VAR
(* ENGINEERING_CONTRACT
 * Parse dotted-decimal IPv4 string to 32-bit network-order UDINT.
 * Input:  ipText (STRING(254)) - dotted-decimal address
 * Output: ipValue (UDINT) - 32-bit value, network byte order; 0 if invalid
 *
 * PUB001: Parse ipText for exactly 4 decimal-digit segments separated by 3 periods
 * PUB002: Each segment value must be 0-255 inclusive
 * PUB003: Network byte order: seg1=MSB<<24, seg2<<16, seg3<<8, seg4=LSB
 * PUB004: Invalid input (wrong count, nondigit, OOR, empty segment) → ipValue=0
 *         Note: Valid address 0.0.0.0 also produces 0 per spec.
 *
 * Contract behavior: Pure combinational, no latches, no state retention.
 * Output ipValue is defined every scan from current ipText.
 *)

ipValue := 0;
tmp_valid := TRUE;

tmp_dot1 := FIND(ipText, '.');
IF tmp_dot1 < 2 OR tmp_dot1 >= LEN(ipText) THEN
    tmp_valid := FALSE;
END_IF

IF tmp_valid THEN
    tmp_dot2 := FIND(MID(ipText, LEN(ipText) - tmp_dot1, tmp_dot1 + 1), '.');
    IF tmp_dot2 < 2 OR tmp_dot2 >= (LEN(ipText) - tmp_dot1) THEN
        tmp_valid := FALSE;
    END_IF;
END_IF

IF tmp_valid THEN
    tmp_dot3 := FIND(MID(ipText, LEN(ipText) - (tmp_dot1 + tmp_dot2), tmp_dot1 + tmp_dot2 + 1), '.');
    IF tmp_dot3 < 2 THEN
        tmp_valid := FALSE;
    END_IF;
END_IF;

IF tmp_valid THEN
    tmp_seg1 := LEFT(ipText, tmp_dot1 - 1);
    tmp_seg2 := MID(ipText, tmp_dot2 - 1, tmp_dot1 + 1);
    tmp_seg3 := MID(ipText, tmp_dot3 - 1, tmp_dot1 + tmp_dot2 + 1);
    tmp_seg4 := MID(ipText, LEN(ipText) - (tmp_dot1 + tmp_dot2 + tmp_dot3), tmp_dot1 + tmp_dot2 + tmp_dot3 + 1);

    // Validate segment 1
    IF LEN(tmp_seg1) < 1 OR LEN(tmp_seg1) > 3 THEN
        tmp_valid := FALSE;
    ELSE
        tmp_val1 := 0;
        FOR tmp_i := 1 TO LEN(tmp_seg1) DO
            tmp_ch := MID(tmp_seg1, 1, tmp_i);
            IF tmp_ch < 48 OR tmp_ch > 57 THEN
                tmp_valid := FALSE;
                EXIT;
            END_IF
            tmp_val1 := tmp_val1 * 10 + TO_UDINT(tmp_ch - 48);
        END_FOR
        IF tmp_val1 > 255 THEN
            tmp_valid := FALSE;
        END_IF
    END_IF

    // Validate segment 2
    IF tmp_valid AND (LEN(tmp_seg2) < 1 OR LEN(tmp_seg2) > 3) THEN
        tmp_valid := FALSE;
    END_IF

    IF tmp_valid THEN
        tmp_val2 := 0;
        FOR tmp_i := 1 TO LEN(tmp_seg2) DO
            tmp_ch := MID(tmp_seg2, 1, tmp_i);
            IF tmp_ch < 48 OR tmp_ch > 57 THEN
                tmp_valid := FALSE;
                EXIT;
            END_IF
            tmp_val2 := tmp_val2 * 10 + TO_UDINT(tmp_ch - 48);
        END_FOR
        IF tmp_val2 > 255 THEN
            tmp_valid := FALSE;
        END_IF
    END_IF

    // Validate segment 3
    IF tmp_valid AND (LEN(tmp_seg3) < 1 OR LEN(tmp_seg3) > 3) THEN
        tmp_valid := FALSE;
    END_IF

    IF tmp_valid THEN
        tmp_val3 := 0;
        FOR tmp_i := 1 TO LEN(tmp_seg3) DO
            tmp_ch := MID(tmp_seg3, 1, tmp_i);
            IF tmp_ch < 48 OR tmp_ch > 57 THEN
                tmp_valid := FALSE;
                EXIT;
            END_IF
            tmp_val3 := tmp_val3 * 10 + TO_UDINT(tmp_ch - 48);
        END_FOR
        IF tmp_val3 > 255 THEN
            tmp_valid := FALSE;
        END_IF
    END_IF

    // Validate segment 4
    IF tmp_valid AND (LEN(tmp_seg4) < 1 OR LEN(tmp_seg4) > 3) THEN
        tmp_valid := FALSE;
    END_IF

    IF tmp_valid THEN
        tmp_val4 := 0;
        FOR tmp_i := 1 TO LEN(tmp_seg4) DO
            tmp_ch := MID(tmp_seg4, 1, tmp_i);
            IF tmp_ch < 48 OR tmp_ch > 57 THEN
                tmp_valid := FALSE;
                EXIT;
            END_IF
            tmp_val4 := tmp_val4 * 10 + TO_UDINT(tmp_ch - 48);
        END_FOR
        IF tmp_val4 > 255 THEN
            tmp_valid := FALSE;
        END_IF
    END_IF
END_IF

IF tmp_valid THEN
    ipValue := SHL(tmp_val1, 24) OR SHL(tmp_val2, 16) OR SHL(tmp_val3, 8) OR tmp_val4;
END_IF

END_FUNCTION_BLOCK
(* CONTRACT_RULES [] *)

(* ---- public-medium-08.raw_candidate_03.st ---- *)
FUNCTION_BLOCK FB_IPv4Parse
VAR_INPUT
    ipText : STRING(254);
END_VAR
VAR_OUTPUT
    ipValue : UDINT;
END_VAR
VAR
    tmp_dot1 : INT;
    tmp_dot2 : INT;
    tmp_dot3 : INT;
    tmp_seg1 : STRING(4);
    tmp_seg2 : STRING(4);
    tmp_seg3 : STRING(4);
    tmp_seg4 : STRING(4);
    tmp_val1 : UDINT;
    tmp_val2 : UDINT;
    tmp_val3 : UDINT;
    tmp_val4 : UDINT;
    tmp_valid : BOOL;
    tmp_i : INT;
    tmp_ch : BYTE;
END_VAR
(* ENGINEERING_CONTRACT
 * Parse dotted-decimal IPv4 string to 32-bit network-order UDINT.
 * Input:  ipText (STRING(254)) - dotted-decimal address
 * Output: ipValue (UDINT) - 32-bit value, network byte order; 0 if invalid
 *
 * PUB001: Parse ipText for exactly 4 decimal-digit segments separated by 3 periods
 * PUB002: Each segment value must be 0-255 inclusive
 * PUB003: Network byte order: seg1=MSB<<24, seg2<<16, seg3<<8, seg4=LSB
 * PUB004: Invalid input (wrong count, nondigit, OOR, empty segment) → ipValue=0
 *         Note: Valid address 0.0.0.0 also produces 0 per spec.
 *
 * Contract behavior: Pure combinational, no latches, no state retention.
 * Output ipValue is defined every scan from current ipText.
 *)

ipValue := 0;
tmp_valid := TRUE;

tmp_dot1 := FIND(ipText, '.');
IF tmp_dot1 < 2 OR tmp_dot1 >= LEN(ipText) THEN
    tmp_valid := FALSE;
END_IF;

IF tmp_valid THEN
    tmp_dot2 := FIND(MID(ipText, LEN(ipText) - tmp_dot1, tmp_dot1 + 1), '.');
    IF tmp_dot2 < 2 OR tmp_dot2 >= (LEN(ipText) - tmp_dot1) THEN
        tmp_valid := FALSE;
    END_IF;
END_IF;

IF tmp_valid THEN
    tmp_dot3 := FIND(MID(ipText, LEN(ipText) - (tmp_dot1 + tmp_dot2), tmp_dot1 + tmp_dot2 + 1), '.');
    IF tmp_dot3 < 2 THEN
        tmp_valid := FALSE;
    END_IF;
END_IF;

IF tmp_valid THEN
    tmp_seg1 := LEFT(ipText, tmp_dot1 - 1);
    tmp_seg2 := MID(ipText, tmp_dot2 - 1, tmp_dot1 + 1);
    tmp_seg3 := MID(ipText, tmp_dot3 - 1, tmp_dot1 + tmp_dot2 + 1);
    tmp_seg4 := MID(ipText, LEN(ipText) - (tmp_dot1 + tmp_dot2 + tmp_dot3), tmp_dot1 + tmp_dot2 + tmp_dot3 + 1);

    // Validate segment 1
    IF LEN(tmp_seg1) < 1 OR LEN(tmp_seg1) > 3 THEN
        tmp_valid := FALSE;
    ELSE
        tmp_val1 := 0;
        FOR tmp_i := 1 TO LEN(tmp_seg1) DO
            tmp_ch := ipText[tmp_i];
            IF tmp_ch < 48 OR tmp_ch > 57 THEN
                tmp_valid := FALSE;
                EXIT;
            END_IF;
            tmp_val1 := tmp_val1 * 10 + TO_UDINT(tmp_ch - 48);
        END_FOR;
        IF tmp_val1 > 255 THEN
            tmp_valid := FALSE;
        END_IF;
    END_IF;

    // Validate segment 2
    IF tmp_valid AND (LEN(tmp_seg2) < 1 OR LEN(tmp_seg2) > 3) THEN
        tmp_valid := FALSE;
    END_IF;

    IF tmp_valid THEN
        tmp_val2 := 0;
        FOR tmp_i := 1 TO LEN(tmp_seg2) DO
            tmp_ch := ipText[tmp_dot1 + tmp_dot2 + tmp_i];
            IF tmp_ch < 48 OR tmp_ch > 57 THEN
                tmp_valid := FALSE;
                EXIT;
            END_IF;
            tmp_val2 := tmp_val2 * 10 + TO_UDINT(tmp_ch - 48);
        END_FOR;
        IF tmp_val2 > 255 THEN
            tmp_valid := FALSE;
        END_IF;
    END_IF;

    // Validate segment 3
    IF tmp_valid AND (LEN(tmp_seg3) < 1 OR LEN(tmp_seg3) > 3) THEN
        tmp_valid := FALSE;
    END_IF;

    IF tmp_valid THEN
        tmp_val3 := 0;
        FOR tmp_i := 1 TO LEN(tmp_seg3) DO
            tmp_ch := ipText[tmp_dot1 + tmp_dot2 + tmp_dot3 + tmp_i];
            IF tmp_ch < 48 OR tmp_ch > 57 THEN
                tmp_valid := FALSE;
                EXIT;
            END_IF;
            tmp_val3 := tmp_val3 * 10 + TO_UDINT(tmp_ch - 48);
        END_FOR;
        IF tmp_val3 > 255 THEN
            tmp_valid := FALSE;
        END_IF;
    END_IF;

    // Validate segment 4
    IF tmp_valid AND (LEN(tmp_seg4) < 1 OR LEN(tmp_seg4) > 3) THEN
        tmp_valid := FALSE;
    END_IF;

    IF tmp_valid THEN
        tmp_val4 := 0;
        FOR tmp_i := 1 TO LEN(tmp_seg4) DO
            tmp_ch := ipText[tmp_dot1 + tmp_dot2 + tmp_dot3 + tmp_i];
            IF tmp_ch < 48 OR tmp_ch > 57 THEN
                tmp_valid := FALSE;
                EXIT;
            END_IF;
            tmp_val4 := tmp_val4 * 10 + TO_UDINT(tmp_ch - 48);
        END_FOR;
        IF tmp_val4 > 255 THEN
            tmp_valid := FALSE;
        END_IF;
    END_IF;
END_IF;

IF tmp_valid THEN
    ipValue := SHL(tmp_val1, 24) OR SHL(tmp_val2, 16) OR SHL(tmp_val3, 8) OR tmp_val4;
END_IF;

END_FUNCTION_BLOCK
(* CONTRACT_RULES [] *)

(* ---- self-easy-01.candidate_01.st ---- *)
(* ENGINEERING_CONTRACT
 * Design table for FB averaging function block:
 *
 * | Output/State  | Activation event             | Retention/hold                  | Explicit reset | Same-scan priority | Units/boundaries      |
 * |---------------|-------------------------------|---------------------------------|----------------|--------------------|-----------------------|
 * | avgOut update | enable AND avgEnable AND      | Hold on: !enable, !avgEnable,   | None stated    | Combinational      | Real, no rounding     |
 * |               | count > 0                     | count <= 0                      |                | override            |                       |
 * | Division      | Only when count > 0 AND       | N/A (blocked)                   | N/A            | N/A                 | Divisor: clamped 1..8 |
 * |               | entering compute branch       |                                 |                |                    |                       |
 * | Sum overflow  | Any valid compute scan        | N/A                             | N/A            | N/A                 | DINT accumulator      |
 *
 * Clause references:
 * - PUB001: enable gate for update
 * - PUB003: count gating, 0..8 range
 * - PUB005: no division by zero
 * - PUB006: count > 8 clamped to 8
 * - PUB007: avgEnable gate
 * - PUB008: DINT sum to avoid overflow
 * - PUB010: REAL output, no rounding
 *
 * Boundary arithmetic:
 * - count = 0: no compute, avgOut held
 * - count = 1..8: compute exactly that many elements
 * - count > 8: compute exactly 8 elements
 * - count < 0: same as count = 0 (held), no negative indexing
 *)

(* CONTRACT_RULES [] *)

FUNCTION_BLOCK FB
VAR_INPUT
    enable    : BOOL;
    values    : ARRAY[1..8] OF INT;
    count     : INT;
    avgEnable : BOOL;
END_VAR

VAR_OUTPUT
    avgOut : REAL;
END_VAR

VAR
    tmp_sum    : DINT;
    tmp_count  : INT;
    i          : INT;
END_VAR

// Compute average only when all gates are active and count is positive
IF enable AND avgEnable AND (count > 0) THEN
    // Clamp effective count to array upper bound
    IF count >= 8 THEN
        tmp_count := 8;
    ELSE
        tmp_count := count;
    END_IF;

    // Accumulate using DINT to prevent INT overflow
    tmp_sum := 0;
    FOR i := 1 TO tmp_count DO
        tmp_sum := tmp_sum + values[i];
    END_FOR;

    // Real division with no rounding
    avgOut := DINT_TO_REAL(tmp_sum) / INT_TO_REAL(tmp_count);
END_IF;
// All other cases: avgOut retains previous value (no assignment)
// Including: !enable, !avgEnable, count <= 0, count < 0
END_FUNCTION_BLOCK

(* ---- self-easy-01.raw_candidate_01.st ---- *)
(* ENGINEERING_CONTRACT
 * Design table for FB averaging function block:
 *
 * | Output/State  | Activation event             | Retention/hold                  | Explicit reset | Same-scan priority | Units/boundaries      |
 * |---------------|-------------------------------|---------------------------------|----------------|--------------------|-----------------------|
 * | avgOut update | enable AND avgEnable AND      | Hold on: !enable, !avgEnable,   | None stated    | Combinational      | Real, no rounding     |
 * |               | count > 0                     | count <= 0                      |                | override            |                       |
 * | Division      | Only when count > 0 AND       | N/A (blocked)                   | N/A            | N/A                 | Divisor: clamped 1..8 |
 * |               | entering compute branch       |                                 |                |                    |                       |
 * | Sum overflow  | Any valid compute scan        | N/A                             | N/A            | N/A                 | DINT accumulator      |
 *
 * Clause references:
 * - PUB001: enable gate for update
 * - PUB003: count gating, 0..8 range
 * - PUB005: no division by zero
 * - PUB006: count > 8 clamped to 8
 * - PUB007: avgEnable gate
 * - PUB008: DINT sum to avoid overflow
 * - PUB010: REAL output, no rounding
 *
 * Boundary arithmetic:
 * - count = 0: no compute, avgOut held
 * - count = 1..8: compute exactly that many elements
 * - count > 8: compute exactly 8 elements
 * - count < 0: same as count = 0 (held), no negative indexing
 *)

(* CONTRACT_RULES [] *)

FUNCTION_BLOCK FB
VAR_INPUT
    enable    : BOOL;
    values    : ARRAY[1..8] OF INT;
    count     : INT;
    avgEnable : BOOL;
END_VAR

VAR_OUTPUT
    avgOut : REAL;
END_VAR

VAR
    tmp_sum    : DINT;
    tmp_count  : INT;
    i          : INT;
END_VAR

// Compute average only when all gates are active and count is positive
IF enable AND avgEnable AND (count > 0) THEN
    // Clamp effective count to array upper bound
    IF count >= 8 THEN
        tmp_count := 8;
    ELSE
        tmp_count := count;
    END_IF;

    // Accumulate using DINT to prevent INT overflow
    tmp_sum := 0;
    FOR i := 1 TO tmp_count DO
        tmp_sum := tmp_sum + values[i];
    END_FOR;

    // Real division with no rounding
    avgOut := DINT_TO_REAL(tmp_sum) / INT_TO_REAL(tmp_count);
END_IF;
// All other cases: avgOut retains previous value (no assignment)
// Including: !enable, !avgEnable, count <= 0, count < 0
END_FUNCTION_BLOCK

(* ---- self-easy-02.candidate_01.st ---- *)
(* CONTRACT_RULES [{"kind":"hold_until_reset","output":"alarmHigh","set_input":"tankLevel","reset_input":"resetBtn"},{"kind":"hold_until_reset","output":"alarmLow","set_input":"tankLevel","reset_input":"resetBtn"}] *)

(* ENGINEERING_CONTRACT
 * Input sampling: tankLevel, inletPermit, resetBtn sampled each scan
 * Output update: all outputs evaluated at end of same scan
 *
 * | Output     | Activation              | Retention                  | Reset/Deactivation           | Priority      |
 * |------------|-------------------------|----------------------------|------------------------------|---------------|
 * | alarmHigh  | tankLevel >= 85.0       | Latched until safe+reset   | rising(resetBtn) & level<85  | Immediate     |
 * | alarmLow   | tankLevel <= 15.0       | Latched until safe+reset   | rising(resetBtn) & level>15  | Immediate     |
 * | pumpRun    | inletPermit & !alarms   | Held while conditions met  | Any alarm active or !permit  | Stop > Start  |
 * | outletValveOpen | !alarmLow           | Open unless low alarm held | alarmLow active closes it    | Inverse of alarmLow |
 *
 * Boundaries: high=85.0, low=15.0 (inclusive thresholds per PUB001/PUB002)
 * Initial state: all outputs FALSE, prevBtn=FALSE
 * Scan behavior: same-scan evaluation of final state, edge detected via prev state
 *)

FUNCTION_BLOCK FB
VAR_INPUT
    tankLevel   : REAL;
    outletFlow  : REAL;
    inletPermit : BOOL;
    resetBtn    : BOOL;
END_VAR
VAR_OUTPUT
    pumpRun         : BOOL;
    alarmHigh       : BOOL;
    alarmLow        : BOOL;
    outletValveOpen : BOOL;
END_VAR
VAR
    prevResetBtn : BOOL := FALSE;
    prevAlarmHigh : BOOL := FALSE;
    prevAlarmLow  : BOOL := FALSE;
    tmpRisingReset : BOOL;
    tmpLevelHigh   : BOOL;
    tmpLevelLow    : BOOL;
END_VAR

    tmpRisingReset := resetBtn AND NOT prevResetBtn;
    tmpLevelHigh := (tankLevel >= 85.0);
    tmpLevelLow  := (tankLevel <= 15.0);

    IF tmpLevelHigh THEN
        alarmHigh := TRUE;
    ELSIF tmpRisingReset AND NOT tmpLevelHigh THEN
        alarmHigh := FALSE;
    END_IF;

    IF tmpLevelLow THEN
        alarmLow := TRUE;
    ELSIF tmpRisingReset AND NOT tmpLevelLow THEN
        alarmLow := FALSE;
    END_IF;

    IF NOT alarmHigh AND NOT alarmLow AND inletPermit THEN
        pumpRun := TRUE;
    ELSE
        pumpRun := FALSE;
    END_IF;

    outletValveOpen := NOT alarmLow;

    prevResetBtn := resetBtn;
    prevAlarmHigh := alarmHigh;
    prevAlarmLow := alarmLow;
END_FUNCTION_BLOCK

(* ---- self-easy-02.raw_candidate_01.st ---- *)
(* CONTRACT_RULES [{"kind":"hold_until_reset","output":"alarmHigh","set_input":"tankLevel","reset_input":"resetBtn"},{"kind":"hold_until_reset","output":"alarmLow","set_input":"tankLevel","reset_input":"resetBtn"}] *)

(* ENGINEERING_CONTRACT
 * Input sampling: tankLevel, inletPermit, resetBtn sampled each scan
 * Output update: all outputs evaluated at end of same scan
 *
 * | Output     | Activation              | Retention                  | Reset/Deactivation           | Priority      |
 * |------------|-------------------------|----------------------------|------------------------------|---------------|
 * | alarmHigh  | tankLevel >= 85.0       | Latched until safe+reset   | rising(resetBtn) & level<85  | Immediate     |
 * | alarmLow   | tankLevel <= 15.0       | Latched until safe+reset   | rising(resetBtn) & level>15  | Immediate     |
 * | pumpRun    | inletPermit & !alarms   | Held while conditions met  | Any alarm active or !permit  | Stop > Start  |
 * | outletValveOpen | !alarmLow           | Open unless low alarm held | alarmLow active closes it    | Inverse of alarmLow |
 *
 * Boundaries: high=85.0, low=15.0 (inclusive thresholds per PUB001/PUB002)
 * Initial state: all outputs FALSE, prevBtn=FALSE
 * Scan behavior: same-scan evaluation of final state, edge detected via prev state
 *)

FUNCTION_BLOCK FB
VAR_INPUT
    tankLevel   : REAL;
    outletFlow  : REAL;
    inletPermit : BOOL;
    resetBtn    : BOOL;
END_VAR
VAR_OUTPUT
    pumpRun         : BOOL;
    alarmHigh       : BOOL;
    alarmLow        : BOOL;
    outletValveOpen : BOOL;
END_VAR
VAR
    prevResetBtn : BOOL := FALSE;
    prevAlarmHigh : BOOL := FALSE;
    prevAlarmLow  : BOOL := FALSE;
    tmpRisingReset : BOOL;
    tmpLevelHigh   : BOOL;
    tmpLevelLow    : BOOL;
END_VAR

    tmpRisingReset := resetBtn AND NOT prevResetBtn;
    tmpLevelHigh := (tankLevel >= 85.0);
    tmpLevelLow  := (tankLevel <= 15.0);

    IF tmpLevelHigh THEN
        alarmHigh := TRUE;
    ELSIF tmpRisingReset AND NOT tmpLevelHigh THEN
        alarmHigh := FALSE;
    END_IF;

    IF tmpLevelLow THEN
        alarmLow := TRUE;
    ELSIF tmpRisingReset AND NOT tmpLevelLow THEN
        alarmLow := FALSE;
    END_IF;

    IF NOT alarmHigh AND NOT alarmLow AND inletPermit THEN
        pumpRun := TRUE;
    ELSE
        pumpRun := FALSE;
    END_IF;

    outletValveOpen := NOT alarmLow;

    prevResetBtn := resetBtn;
    prevAlarmHigh := alarmHigh;
    prevAlarmLow := alarmLow;
END_FUNCTION_BLOCK

(* ---- self-hard-01.candidate_01.st ---- *)
FUNCTION_BLOCK FB
VAR_INPUT
    flowLow   : BOOL;
    ackBtn    : BOOL;
    sensorOK  : BOOL;
END_VAR
VAR_OUTPUT
    alarmActive : BOOL;
    alarmAcked  : BOOL;
    highHigh    : BOOL;
END_VAR
VAR
    prev_flowLow  : BOOL := FALSE;
    prev_alarmActive : BOOL := FALSE;
    prev_alarmAcked  : BOOL := FALSE;
END_VAR
VAR_TEMP
    ackRising : BOOL;
END_VAR
(* ENGINEERING_CONTRACT
   ISA-18.2 four-state alarm (unack-active / unack-cleared / acked-active / acked-cleared):
   ┌──────────────────┬───────────────┬──────────────────────────────────────────────┐
   │ Output / State   │ Activation    │ Retention / Reset / Deactivation              │
   ├──────────────────┼───────────────┼──────────────────────────────────────────────┤
   │ alarmActive      │ flowLow rising│ Held until condition cleared AND alarmAcked   │
   │                  │ edge          │ (no self-clear without explicit ack)         │
   ├──────────────────┼───────────────┼──────────────────────────────────────────────┤
   │ alarmAcked       │ 1) ackBtn     │ Held across scans; reset only when acked-btn │
   │                  │    rising edge│    pressed while condition gone (clears both)│
   │                  │ 2) condition  │                                              │
   │                  │    cleared    │                                              │
   │                  │    (prev unack│                                              │
   │                  │    active)    │                                              │
   ├──────────────────┼───────────────┼──────────────────────────────────────────────┤
   │ highHigh         │ sensorOK=FALSE│ Auto-cleared when sensorOK returns TRUE      │
   │                  │ (same scan)   │ (independent, never inhibits low alarm)     │
   └──────────────────┴───────────────┴──────────────────────────────────────────────┘
   Boundaries:
     - alarmActive retained across scans when !alarmAcked (PUB001/PUB002/PUB005)
     - highHigh = NOT sensorOK  (PUB004/PUB016)
     - ackBtn rising-edge only; same-scan evaluation (PUB006/PUB007/PUB014)
     - No timers or hidden state; all VAR static (PUB008)
   Supported formal properties:
     [S1] G(flowLow & ackBtn -> alarmActive)
     [S2] G(alarmActive & !alarmAcked & X(flowLow) -> X(alarmActive))
     [S3] G(!sensorOK -> highHigh)
     [S4] G(rising(ackBtn) & flowLow -> alarmAcked)
     [S5] G(highHigh <-> !sensorOK)
     [S6] alarmActive FSM (see state table above)
     [S7] alarmAcked FSM (see state table above)
*)
BEGIN
    (* Rising-edge detection *)
    ackRising := ackBtn AND NOT prev_alarmActive; (* reuse prev_alarmActive as prev_ackBtn *)

    (* ── High-priority alarm: sensor wire-break ── *)
    highHigh := NOT sensorOK;  (* PUB004/PUB016, PUB034: auto-clear when OK *)

    (* ── Four-state low-priority alarm ── *)

    (* Condition gone transitions *)
    IF flowLow THEN
        (* Condition still present *)
        alarmActive := TRUE;
        IF ackRising THEN
            alarmAcked := TRUE;  (* acked while condition present: acked-active *)
        END_IF;
    ELSE
        (* Condition currently gone *)
        IF prev_flowLow THEN
            (* Just-cleared edge: alarm can't vanish unacknowledged *)
            IF alarmActive AND NOT alarmAcked THEN
                alarmAcked := TRUE;   (* unack-active → acked-cleared *)
            END_IF;
            (* acked-cleared stays active until user presses ack *)
            IF alarmActive AND alarmAcked THEN
                (* stay acked-cleared; handled below after ack check *)
            END_IF;
        END_IF;

        (* Transition out of acked-cleared on explicit acknowledge *)
        IF alarmActive AND alarmAcked AND ackRising THEN
            alarmActive := FALSE;
            alarmAcked  := FALSE;
        END_IF;

        (* No active alarm and not just cleared → cleared state *)
        IF NOT alarmActive THEN
            alarmAcked := FALSE;
        END_IF;
    END_IF;

    (* Persist alarmActive when condition present but not yet acked *)
    IF flowLow AND prev_flowLow AND alarmActive AND NOT alarmAcked THEN
        alarmActive := TRUE;   (* hold unack-active across scans *)
    END_IF;

    (* Shift-register for next scan *)
    prev_flowLow     := flowLow;
    prev_alarmActive := alarmActive;
    prev_alarmAcked  := alarmAcked;
    (* reuse: prev_alarmActive used as prev_ackBtn above via ackRising *)
END_FUNCTION_BLOCK

(* ---- self-hard-01.candidate_02.st ---- *)
FUNCTION_BLOCK FB
VAR_INPUT
    flowLow   : BOOL;
    ackBtn    : BOOL;
    sensorOK  : BOOL;
END_VAR
VAR_OUTPUT
    alarmActive : BOOL;
    alarmAcked  : BOOL;
    highHigh    : BOOL;
END_VAR
VAR
    prev_flowLow  : BOOL := FALSE;
    prev_ackBtn   : BOOL := FALSE;
    prev_alarmActive : BOOL := FALSE;
    prev_alarmAcked  : BOOL := FALSE;
END_VAR
VAR_TEMP
    ackRising : BOOL;
END_VAR
(* ENGINEERING_CONTRACT
   ISA-18.2 four-state alarm (unack-active / unack-cleared / acked-active / acked-cleared):
   ┌──────────────────┬───────────────┬──────────────────────────────────────────────┐
   │ Output / State   │ Activation    │ Retention / Reset / Deactivation              │
   ├──────────────────┼───────────────┼──────────────────────────────────────────────┤
   │ alarmActive      │ flowLow rising│ Held until condition cleared AND alarmAcked   │
   │                  │ edge          │ (no self-clear without explicit ack)         │
   ├──────────────────┼───────────────┼──────────────────────────────────────────────┤
   │ alarmAcked       │ 1) ackBtn     │ Held across scans; reset only when acked-btn │
   │                  │    rising edge│    pressed while condition gone (clears both)│
   │                  │ 2) condition  │                                              │
   │                  │    cleared    │                                              │
   │                  │    (prev unack│                                              │
   │                  │    active)    │                                              │
   ├──────────────────┼───────────────┼──────────────────────────────────────────────┤
   │ highHigh         │ sensorOK=FALSE│ Auto-cleared when sensorOK returns TRUE      │
   │                  │ (same scan)   │ (independent, never inhibits low alarm)     │
   └──────────────────┴───────────────┴──────────────────────────────────────────────┘
   Boundaries:
     - alarmActive retained across scans when !alarmAcked (PUB001/PUB002/PUB005)
     - highHigh = NOT sensorOK  (PUB004/PUB016)
     - ackBtn rising-edge only; same-scan evaluation (PUB006/PUB007/PUB014)
     - No timers or hidden state; all VAR static (PUB008)
   Supported formal properties:
     [S1] G(flowLow & ackBtn -> alarmActive)
     [S2] G(alarmActive & !alarmAcked & X(flowLow) -> X(alarmActive))
     [S3] G(!sensorOK -> highHigh)
     [S4] G(rising(ackBtn) & flowLow -> alarmAcked)
     [S5] G(highHigh <-> !sensorOK)
     [S6] alarmActive FSM (see state table above)
     [S7] alarmAcked FSM (see state table above)
*)
    (* Rising-edge detection *)
    ackRising := ackBtn AND NOT prev_ackBtn;

    (* ── High-priority alarm: sensor wire-break ── *)
    highHigh := NOT sensorOK;  (* PUB004/PUB016, PUB034: auto-clear when OK *)

    (* ── Four-state low-priority alarm ── *)

    (* Condition gone transitions *)
    IF flowLow THEN
        (* Condition still present *)
        alarmActive := TRUE;
        IF ackRising THEN
            alarmAcked := TRUE;  (* acked while condition present: acked-active *)
        END_IF;
    ELSE
        (* Condition currently gone *)
        IF prev_flowLow THEN
            (* Just-cleared edge: alarm can't vanish unacknowledged *)
            IF alarmActive AND NOT alarmAcked THEN
                alarmAcked := TRUE;   (* unack-active → acked-cleared *)
            END_IF;
            (* acked-cleared stays active until user presses ack *)
            IF alarmActive AND alarmAcked THEN
                (* stay acked-cleared; handled below after ack check *)
            END_IF;
        END_IF;

        (* Transition out of acked-cleared on explicit acknowledge *)
        IF alarmActive AND alarmAcked AND ackRising THEN
            alarmActive := FALSE;
            alarmAcked  := FALSE;
        END_IF;

        (* No active alarm and not just cleared → cleared state *)
        IF NOT alarmActive THEN
            alarmAcked := FALSE;
        END_IF;
    END_IF;

    (* Persist alarmActive when condition present but not yet acked *)
    IF flowLow AND prev_flowLow AND alarmActive AND NOT alarmAcked THEN
        alarmActive := TRUE;   (* hold unack-active across scans *)
    END_IF;

    (* Shift-register for next scan *)
    prev_flowLow     := flowLow;
    prev_ackBtn      := ackBtn;
    prev_alarmActive := alarmActive;
    prev_alarmAcked  := alarmAcked;
END_FUNCTION_BLOCK

(* ---- self-hard-01.candidate_03.st ---- *)
FUNCTION_BLOCK FB
VAR_INPUT
    flowLow   : BOOL;
    ackBtn    : BOOL;
    sensorOK  : BOOL;
END_VAR
VAR_OUTPUT
    alarmActive : BOOL;
    alarmAcked  : BOOL;
    highHigh    : BOOL;
END_VAR
VAR
    prev_flowLow  : BOOL := FALSE;
    prev_ackBtn   : BOOL := FALSE;
    prev_alarmActive : BOOL := FALSE;
    prev_alarmAcked  : BOOL := FALSE;
END_VAR
VAR_TEMP
    ackRising : BOOL;
END_VAR
(* ENGINEERING_CONTRACT
   ISA-18.2 four-state alarm (unack-active / unack-cleared / acked-active / acked-cleared):
   ┌──────────────────┬───────────────┬──────────────────────────────────────────────┐
   │ Output / State   │ Activation    │ Retention / Reset / Deactivation              │
   ├──────────────────┼───────────────┼──────────────────────────────────────────────┤
   │ alarmActive      │ flowLow rising│ Held until condition cleared AND alarmAcked   │
   │                  │ edge          │ (no self-clear without explicit ack)         │
   ├──────────────────┼───────────────┼──────────────────────────────────────────────┤
   │ alarmAcked       │ 1) ackBtn     │ Held across scans; reset only when acked-btn │
   │                  │    rising edge│    pressed while condition gone (clears both)│
   │                  │ 2) condition  │                                              │
   │                  │    cleared    │                                              │
   │                  │    (prev unack│                                              │
   │                  │    active)    │                                              │
   ├──────────────────┼───────────────┼──────────────────────────────────────────────┤
   │ highHigh         │ sensorOK=FALSE│ Auto-cleared when sensorOK returns TRUE      │
   │                  │ (same scan)   │ (independent, never inhibits low alarm)     │
   └──────────────────┴───────────────┴──────────────────────────────────────────────┘
   Boundaries:
     - alarmActive retained across scans when !alarmAcked (PUB001/PUB002/PUB005)
     - highHigh = NOT sensorOK  (PUB004/PUB016)
     - ackBtn rising-edge only; same-scan evaluation (PUB006/PUB007/PUB014)
     - No timers or hidden state; all VAR static (PUB008)
   Supported formal properties:
     [S1] G(flowLow & ackBtn -> alarmActive)
     [S2] G(alarmActive & !alarmAcked & X(flowLow) -> X(alarmActive))
     [S3] G(!sensorOK -> highHigh)
     [S4] G(rising(ackBtn) & flowLow -> alarmAcked)
     [S5] G(highHigh <-> !sensorOK)
     [S6] alarmActive FSM (see state table above)
     [S7] alarmAcked FSM (see state table above)
*)
    ackRising := ackBtn AND NOT prev_ackBtn;

    (* ── High-priority alarm: sensor wire-break ── *)
    highHigh := NOT sensorOK;  (* PUB004/PUB016, PUB034: auto-clear when OK *)

    (* ── Four-state low-priority alarm ── *)

    (* Condition gone transitions *)
    IF flowLow THEN
        (* Condition still present *)
        alarmActive := TRUE;
        IF ackRising THEN
            alarmAcked := TRUE;  (* acked while condition present: acked-active *)
        END_IF;
    ELSE
        (* Condition currently gone *)
        IF prev_flowLow THEN
            (* Just-cleared edge: alarm can't vanish unacknowledged *)
            IF alarmActive AND NOT alarmAcked THEN
                alarmAcked := TRUE;   (* unack-active → acked-cleared *)
            END_IF;
            (* acked-cleared stays active until user presses ack *)
            IF alarmActive AND alarmAcked THEN
                (* stay acked-cleared; handled below after ack check *)
            END_IF;
        END_IF;

        (* Transition out of acked-cleared on explicit acknowledge *)
        IF alarmActive AND alarmAcked AND ackRising THEN
            alarmActive := FALSE;
            alarmAcked  := FALSE;
        END_IF;

        (* No active alarm and not just cleared → cleared state *)
        IF NOT alarmActive THEN
            alarmAcked := FALSE;
        END_IF;
    END_IF;

    (* Persist alarmActive when condition present but not yet acked *)
    IF flowLow AND prev_flowLow AND alarmActive AND NOT alarmAcked THEN
        alarmActive := TRUE;   (* hold unack-active across scans *)
    END_IF;

    (* Shift-register for next scan *)
    prev_flowLow     := flowLow;
    prev_ackBtn      := ackBtn;
    prev_alarmActive := alarmActive;
    prev_alarmAcked  := alarmAcked;
END_FUNCTION_BLOCK

(* ---- self-hard-01.patch_base_02.st ---- *)
FUNCTION_BLOCK FB
VAR_INPUT
    flowLow   : BOOL;
    ackBtn    : BOOL;
    sensorOK  : BOOL;
END_VAR
VAR_OUTPUT
    alarmActive : BOOL;
    alarmAcked  : BOOL;
    highHigh    : BOOL;
END_VAR
VAR
    prev_flowLow  : BOOL := FALSE;
    prev_alarmActive : BOOL := FALSE;
    prev_alarmAcked  : BOOL := FALSE;
END_VAR
VAR_TEMP
    ackRising : BOOL;
END_VAR
(* ENGINEERING_CONTRACT
   ISA-18.2 four-state alarm (unack-active / unack-cleared / acked-active / acked-cleared):
   ┌──────────────────┬───────────────┬──────────────────────────────────────────────┐
   │ Output / State   │ Activation    │ Retention / Reset / Deactivation              │
   ├──────────────────┼───────────────┼──────────────────────────────────────────────┤
   │ alarmActive      │ flowLow rising│ Held until condition cleared AND alarmAcked   │
   │                  │ edge          │ (no self-clear without explicit ack)         │
   ├──────────────────┼───────────────┼──────────────────────────────────────────────┤
   │ alarmAcked       │ 1) ackBtn     │ Held across scans; reset only when acked-btn │
   │                  │    rising edge│    pressed while condition gone (clears both)│
   │                  │ 2) condition  │                                              │
   │                  │    cleared    │                                              │
   │                  │    (prev unack│                                              │
   │                  │    active)    │                                              │
   ├──────────────────┼───────────────┼──────────────────────────────────────────────┤
   │ highHigh         │ sensorOK=FALSE│ Auto-cleared when sensorOK returns TRUE      │
   │                  │ (same scan)   │ (independent, never inhibits low alarm)     │
   └──────────────────┴───────────────┴──────────────────────────────────────────────┘
   Boundaries:
     - alarmActive retained across scans when !alarmAcked (PUB001/PUB002/PUB005)
     - highHigh = NOT sensorOK  (PUB004/PUB016)
     - ackBtn rising-edge only; same-scan evaluation (PUB006/PUB007/PUB014)
     - No timers or hidden state; all VAR static (PUB008)
   Supported formal properties:
     [S1] G(flowLow & ackBtn -> alarmActive)
     [S2] G(alarmActive & !alarmAcked & X(flowLow) -> X(alarmActive))
     [S3] G(!sensorOK -> highHigh)
     [S4] G(rising(ackBtn) & flowLow -> alarmAcked)
     [S5] G(highHigh <-> !sensorOK)
     [S6] alarmActive FSM (see state table above)
     [S7] alarmAcked FSM (see state table above)
*)
BEGIN
    (* Rising-edge detection *)
    ackRising := ackBtn AND NOT prev_alarmActive; (* reuse prev_alarmActive as prev_ackBtn *)

    (* ── High-priority alarm: sensor wire-break ── *)
    highHigh := NOT sensorOK;  (* PUB004/PUB016, PUB034: auto-clear when OK *)

    (* ── Four-state low-priority alarm ── *)

    (* Condition gone transitions *)
    IF flowLow THEN
        (* Condition still present *)
        alarmActive := TRUE;
        IF ackRising THEN
            alarmAcked := TRUE;  (* acked while condition present: acked-active *)
        END_IF;
    ELSE
        (* Condition currently gone *)
        IF prev_flowLow THEN
            (* Just-cleared edge: alarm can't vanish unacknowledged *)
            IF alarmActive AND NOT alarmAcked THEN
                alarmAcked := TRUE;   (* unack-active → acked-cleared *)
            END_IF;
            (* acked-cleared stays active until user presses ack *)
            IF alarmActive AND alarmAcked THEN
                (* stay acked-cleared; handled below after ack check *)
            END_IF;
        END_IF;

        (* Transition out of acked-cleared on explicit acknowledge *)
        IF alarmActive AND alarmAcked AND ackRising THEN
            alarmActive := FALSE;
            alarmAcked  := FALSE;
        END_IF;

        (* No active alarm and not just cleared → cleared state *)
        IF NOT alarmActive THEN
            alarmAcked := FALSE;
        END_IF;
    END_IF;

    (* Persist alarmActive when condition present but not yet acked *)
    IF flowLow AND prev_flowLow AND alarmActive AND NOT alarmAcked THEN
        alarmActive := TRUE;   (* hold unack-active across scans *)
    END_IF;

    (* Shift-register for next scan *)
    prev_flowLow     := flowLow;
    prev_alarmActive := alarmActive;
    prev_alarmAcked  := alarmAcked;
    (* reuse: prev_alarmActive used as prev_ackBtn above via ackRising *)
END_FUNCTION_BLOCK

(* ---- self-hard-01.patch_base_03.st ---- *)
FUNCTION_BLOCK FB
VAR_INPUT
    flowLow   : BOOL;
    ackBtn    : BOOL;
    sensorOK  : BOOL;
END_VAR
VAR_OUTPUT
    alarmActive : BOOL;
    alarmAcked  : BOOL;
    highHigh    : BOOL;
END_VAR
VAR
    prev_flowLow  : BOOL := FALSE;
    prev_ackBtn   : BOOL := FALSE;
    prev_alarmActive : BOOL := FALSE;
    prev_alarmAcked  : BOOL := FALSE;
END_VAR
VAR_TEMP
    ackRising : BOOL;
END_VAR
(* ENGINEERING_CONTRACT
   ISA-18.2 four-state alarm (unack-active / unack-cleared / acked-active / acked-cleared):
   ┌──────────────────┬───────────────┬──────────────────────────────────────────────┐
   │ Output / State   │ Activation    │ Retention / Reset / Deactivation              │
   ├──────────────────┼───────────────┼──────────────────────────────────────────────┤
   │ alarmActive      │ flowLow rising│ Held until condition cleared AND alarmAcked   │
   │                  │ edge          │ (no self-clear without explicit ack)         │
   ├──────────────────┼───────────────┼──────────────────────────────────────────────┤
   │ alarmAcked       │ 1) ackBtn     │ Held across scans; reset only when acked-btn │
   │                  │    rising edge│    pressed while condition gone (clears both)│
   │                  │ 2) condition  │                                              │
   │                  │    cleared    │                                              │
   │                  │    (prev unack│                                              │
   │                  │    active)    │                                              │
   ├──────────────────┼───────────────┼──────────────────────────────────────────────┤
   │ highHigh         │ sensorOK=FALSE│ Auto-cleared when sensorOK returns TRUE      │
   │                  │ (same scan)   │ (independent, never inhibits low alarm)     │
   └──────────────────┴───────────────┴──────────────────────────────────────────────┘
   Boundaries:
     - alarmActive retained across scans when !alarmAcked (PUB001/PUB002/PUB005)
     - highHigh = NOT sensorOK  (PUB004/PUB016)
     - ackBtn rising-edge only; same-scan evaluation (PUB006/PUB007/PUB014)
     - No timers or hidden state; all VAR static (PUB008)
   Supported formal properties:
     [S1] G(flowLow & ackBtn -> alarmActive)
     [S2] G(alarmActive & !alarmAcked & X(flowLow) -> X(alarmActive))
     [S3] G(!sensorOK -> highHigh)
     [S4] G(rising(ackBtn) & flowLow -> alarmAcked)
     [S5] G(highHigh <-> !sensorOK)
     [S6] alarmActive FSM (see state table above)
     [S7] alarmAcked FSM (see state table above)
*)
    (* Rising-edge detection *)
    ackRising := ackBtn AND NOT prev_ackBtn;

    (* ── High-priority alarm: sensor wire-break ── *)
    highHigh := NOT sensorOK;  (* PUB004/PUB016, PUB034: auto-clear when OK *)

    (* ── Four-state low-priority alarm ── *)

    (* Condition gone transitions *)
    IF flowLow THEN
        (* Condition still present *)
        alarmActive := TRUE;
        IF ackRising THEN
            alarmAcked := TRUE;  (* acked while condition present: acked-active *)
        END_IF;
    ELSE
        (* Condition currently gone *)
        IF prev_flowLow THEN
            (* Just-cleared edge: alarm can't vanish unacknowledged *)
            IF alarmActive AND NOT alarmAcked THEN
                alarmAcked := TRUE;   (* unack-active → acked-cleared *)
            END_IF;
            (* acked-cleared stays active until user presses ack *)
            IF alarmActive AND alarmAcked THEN
                (* stay acked-cleared; handled below after ack check *)
            END_IF;
        END_IF;

        (* Transition out of acked-cleared on explicit acknowledge *)
        IF alarmActive AND alarmAcked AND ackRising THEN
            alarmActive := FALSE;
            alarmAcked  := FALSE;
        END_IF;

        (* No active alarm and not just cleared → cleared state *)
        IF NOT alarmActive THEN
            alarmAcked := FALSE;
        END_IF;
    END_IF;

    (* Persist alarmActive when condition present but not yet acked *)
    IF flowLow AND prev_flowLow AND alarmActive AND NOT alarmAcked THEN
        alarmActive := TRUE;   (* hold unack-active across scans *)
    END_IF;

    (* Shift-register for next scan *)
    prev_flowLow     := flowLow;
    prev_ackBtn      := ackBtn;
    prev_alarmActive := alarmActive;
    prev_alarmAcked  := alarmAcked;
END_FUNCTION_BLOCK

(* ---- self-hard-01.patch_base_04.st ---- *)
FUNCTION_BLOCK FB
VAR_INPUT
    flowLow   : BOOL;
    ackBtn    : BOOL;
    sensorOK  : BOOL;
END_VAR
VAR_OUTPUT
    alarmActive : BOOL;
    alarmAcked  : BOOL;
    highHigh    : BOOL;
END_VAR
VAR
    prev_flowLow  : BOOL := FALSE;
    prev_ackBtn   : BOOL := FALSE;
    prev_alarmActive : BOOL := FALSE;
    prev_alarmAcked  : BOOL := FALSE;
END_VAR
VAR_TEMP
    ackRising : BOOL;
END_VAR
(* ENGINEERING_CONTRACT
   ISA-18.2 four-state alarm (unack-active / unack-cleared / acked-active / acked-cleared):
   ┌──────────────────┬───────────────┬──────────────────────────────────────────────┐
   │ Output / State   │ Activation    │ Retention / Reset / Deactivation              │
   ├──────────────────┼───────────────┼──────────────────────────────────────────────┤
   │ alarmActive      │ flowLow rising│ Held until condition cleared AND alarmAcked   │
   │                  │ edge          │ (no self-clear without explicit ack)         │
   ├──────────────────┼───────────────┼──────────────────────────────────────────────┤
   │ alarmAcked       │ 1) ackBtn     │ Held across scans; reset only when acked-btn │
   │                  │    rising edge│    pressed while condition gone (clears both)│
   │                  │ 2) condition  │                                              │
   │                  │    cleared    │                                              │
   │                  │    (prev unack│                                              │
   │                  │    active)    │                                              │
   ├──────────────────┼───────────────┼──────────────────────────────────────────────┤
   │ highHigh         │ sensorOK=FALSE│ Auto-cleared when sensorOK returns TRUE      │
   │                  │ (same scan)   │ (independent, never inhibits low alarm)     │
   └──────────────────┴───────────────┴──────────────────────────────────────────────┘
   Boundaries:
     - alarmActive retained across scans when !alarmAcked (PUB001/PUB002/PUB005)
     - highHigh = NOT sensorOK  (PUB004/PUB016)
     - ackBtn rising-edge only; same-scan evaluation (PUB006/PUB007/PUB014)
     - No timers or hidden state; all VAR static (PUB008)
   Supported formal properties:
     [S1] G(flowLow & ackBtn -> alarmActive)
     [S2] G(alarmActive & !alarmAcked & X(flowLow) -> X(alarmActive))
     [S3] G(!sensorOK -> highHigh)
     [S4] G(rising(ackBtn) & flowLow -> alarmAcked)
     [S5] G(highHigh <-> !sensorOK)
     [S6] alarmActive FSM (see state table above)
     [S7] alarmAcked FSM (see state table above)
*)
    ackRising := ackBtn AND NOT prev_ackBtn;

    (* ── High-priority alarm: sensor wire-break ── *)
    highHigh := NOT sensorOK;  (* PUB004/PUB016, PUB034: auto-clear when OK *)

    (* ── Four-state low-priority alarm ── *)

    (* Condition gone transitions *)
    IF flowLow THEN
        (* Condition still present *)
        alarmActive := TRUE;
        IF ackRising THEN
            alarmAcked := TRUE;  (* acked while condition present: acked-active *)
        END_IF;
    ELSE
        (* Condition currently gone *)
        IF prev_flowLow THEN
            (* Just-cleared edge: alarm can't vanish unacknowledged *)
            IF alarmActive AND NOT alarmAcked THEN
                alarmAcked := TRUE;   (* unack-active → acked-cleared *)
            END_IF;
            (* acked-cleared stays active until user presses ack *)
            IF alarmActive AND alarmAcked THEN
                (* stay acked-cleared; handled below after ack check *)
            END_IF;
        END_IF;

        (* Transition out of acked-cleared on explicit acknowledge *)
        IF alarmActive AND alarmAcked AND ackRising THEN
            alarmActive := FALSE;
            alarmAcked  := FALSE;
        END_IF;

        (* No active alarm and not just cleared → cleared state *)
        IF NOT alarmActive THEN
            alarmAcked := FALSE;
        END_IF;
    END_IF;

    (* Persist alarmActive when condition present but not yet acked *)
    IF flowLow AND prev_flowLow AND alarmActive AND NOT alarmAcked THEN
        alarmActive := TRUE;   (* hold unack-active across scans *)
    END_IF;

    (* Shift-register for next scan *)
    prev_flowLow     := flowLow;
    prev_ackBtn      := ackBtn;
    prev_alarmActive := alarmActive;
    prev_alarmAcked  := alarmAcked;
END_FUNCTION_BLOCK

(* ---- self-hard-01.raw_candidate_01.st ---- *)
FUNCTION_BLOCK FB
VAR_INPUT
    flowLow   : BOOL;
    ackBtn    : BOOL;
    sensorOK  : BOOL;
END_VAR
VAR_OUTPUT
    alarmActive : BOOL;
    alarmAcked  : BOOL;
    highHigh    : BOOL;
END_VAR
VAR
    prev_flowLow  : BOOL := FALSE;
    prev_alarmActive : BOOL := FALSE;
    prev_alarmAcked  : BOOL := FALSE;
END_VAR
VAR_TEMP
    ackRising : BOOL;
END_VAR
(* ENGINEERING_CONTRACT
   ISA-18.2 four-state alarm (unack-active / unack-cleared / acked-active / acked-cleared):
   ┌──────────────────┬───────────────┬──────────────────────────────────────────────┐
   │ Output / State   │ Activation    │ Retention / Reset / Deactivation              │
   ├──────────────────┼───────────────┼──────────────────────────────────────────────┤
   │ alarmActive      │ flowLow rising│ Held until condition cleared AND alarmAcked   │
   │                  │ edge          │ (no self-clear without explicit ack)         │
   ├──────────────────┼───────────────┼──────────────────────────────────────────────┤
   │ alarmAcked       │ 1) ackBtn     │ Held across scans; reset only when acked-btn │
   │                  │    rising edge│    pressed while condition gone (clears both)│
   │                  │ 2) condition  │                                              │
   │                  │    cleared    │                                              │
   │                  │    (prev unack│                                              │
   │                  │    active)    │                                              │
   ├──────────────────┼───────────────┼──────────────────────────────────────────────┤
   │ highHigh         │ sensorOK=FALSE│ Auto-cleared when sensorOK returns TRUE      │
   │                  │ (same scan)   │ (independent, never inhibits low alarm)     │
   └──────────────────┴───────────────┴──────────────────────────────────────────────┘
   Boundaries:
     - alarmActive retained across scans when !alarmAcked (PUB001/PUB002/PUB005)
     - highHigh = NOT sensorOK  (PUB004/PUB016)
     - ackBtn rising-edge only; same-scan evaluation (PUB006/PUB007/PUB014)
     - No timers or hidden state; all VAR static (PUB008)
   Supported formal properties:
     [S1] G(flowLow & ackBtn -> alarmActive)
     [S2] G(alarmActive & !alarmAcked & X(flowLow) -> X(alarmActive))
     [S3] G(!sensorOK -> highHigh)
     [S4] G(rising(ackBtn) & flowLow -> alarmAcked)
     [S5] G(highHigh <-> !sensorOK)
     [S6] alarmActive FSM (see state table above)
     [S7] alarmAcked FSM (see state table above)
*)
BEGIN
    (* Rising-edge detection *)
    ackRising := ackBtn AND NOT prev_alarmActive; (* reuse prev_alarmActive as prev_ackBtn *)

    (* ── High-priority alarm: sensor wire-break ── *)
    highHigh := NOT sensorOK;  (* PUB004/PUB016, PUB034: auto-clear when OK *)

    (* ── Four-state low-priority alarm ── *)

    (* Condition gone transitions *)
    IF flowLow THEN
        (* Condition still present *)
        alarmActive := TRUE;
        IF ackRising THEN
            alarmAcked := TRUE;  (* acked while condition present: acked-active *)
        END_IF
    ELSE
        (* Condition currently gone *)
        IF prev_flowLow THEN
            (* Just-cleared edge: alarm can't vanish unacknowledged *)
            IF alarmActive AND NOT alarmAcked THEN
                alarmAcked := TRUE;   (* unack-active → acked-cleared *)
            END_IF;
            (* acked-cleared stays active until user presses ack *)
            IF alarmActive AND alarmAcked THEN
                (* stay acked-cleared; handled below after ack check *)
            END_IF;
        END_IF;

        (* Transition out of acked-cleared on explicit acknowledge *)
        IF alarmActive AND alarmAcked AND ackRising THEN
            alarmActive := FALSE;
            alarmAcked  := FALSE;
        END_IF;

        (* No active alarm and not just cleared → cleared state *)
        IF NOT alarmActive THEN
            alarmAcked := FALSE;
        END_IF;
    END_IF;

    (* Persist alarmActive when condition present but not yet acked *)
    IF flowLow AND prev_flowLow AND alarmActive AND NOT alarmAcked THEN
        alarmActive := TRUE;   (* hold unack-active across scans *)
    END_IF;

    (* Shift-register for next scan *)
    prev_flowLow     := flowLow;
    prev_alarmActive := alarmActive;
    prev_alarmAcked  := alarmAcked;
    (* reuse: prev_alarmActive used as prev_ackBtn above via ackRising *)
END_FUNCTION_BLOCK
